Universal Robots URScript: test_first_drawing_6_min3.script

def Machining1():
  # Default parameters:
  global speed_ms = 0.3
  global speed_rads = 0.75
  global accel_mss = 3
  global accel_radss = 1.2
  global blend_radius_m = 0.001

  # Add subprograms here
  # Start of main program
  # Program generated by RoboDK v5.6.5 for UR10e on 02/02/2024 17:04:00
  # Using nominal kinematics.
  blend_radius_m = 0.001
  speed_ms = 1.000
  # set_reference(p[0.133734, -0.230000, -0.014586, 0.000000, 0.000000, 0.000000])
  set_tcp(p[0.000000, 0.000000, 0.252000, 0.000000, 0.000000, 0.000000])
  # Show Tool
  movej([-0.330517, -0.653342, -2.600682, -1.458365, 1.570796, 1.240279],accel_radss,speed_rads,0,blend_radius_m)
  movel([-0.330517, -0.653342, -2.600682, -1.458365, 1.570796, 1.240279],accel_mss,speed_ms,0,blend_radius_m)
  # Splitting Linear movement in 6 (instruction 7: MoveL 3)
  movel([-0.330517, -0.660366, -2.629096, -1.422927, 1.570796, 1.240279],accel_mss,speed_ms,0,blend_radius_m)
  movel([-0.330517, -0.669810, -2.657315, -1.385264, 1.570796, 1.240279],accel_mss,speed_ms,0,blend_radius_m)
  movel([-0.330517, -0.682072, -2.685333, -1.344984, 1.570796, 1.240279],accel_mss,speed_ms,0,blend_radius_m)
  movel([-0.330517, -0.697642, -2.713136, -1.301610, 1.570796, 1.240279],accel_mss,speed_ms,0,blend_radius_m)
  movel([-0.330517, -0.717128, -2.740708, -1.254553, 1.570796, 1.240279],accel_mss,speed_ms,0,blend_radius_m)
  movel([-0.330517, -0.741290, -2.768022, -1.203077, 1.570796, 1.240279],accel_mss,speed_ms,0,blend_radius_m)
  movel([-0.330517, -0.741290, -2.768022, -1.203077, 1.570796, 1.240279],accel_mss,speed_ms,0,blend_radius_m)
  speed_ms = 1.000
  movel([-0.330517, -0.741290, -2.768022, -1.203077, 1.570796, 1.240279],accel_mss,speed_ms,0,blend_radius_m)
  movel([-0.330517, -0.741290, -2.768022, -1.203077, 1.570796, 1.240279],accel_mss,speed_ms,0,blend_radius_m)
  movel([-0.330517, -0.741290, -2.768022, -1.203077, 1.570796, 1.240279],accel_mss,speed_ms,0,blend_radius_m)
  speed_ms = 0.005
  movel([-0.330517, -0.712884, -2.735213, -1.264292, 1.570796, 1.240279],accel_mss,speed_ms,0,blend_radius_m)
  speed_ms = 1.000
  movel([-0.330517, -0.741290, -2.768022, -1.203077, 1.570796, 1.240279],accel_mss,speed_ms,0,blend_radius_m)
  speed_ms = 0.040
  movel([-0.330517, -0.741290, -2.768022, -1.203077, 1.570796, 1.240279],accel_mss,speed_ms,0,blend_radius_m)
  speed_ms = 1.000
  movel([-0.330517, -0.741290, -2.768022, -1.203077, 1.570796, 1.240279],accel_mss,speed_ms,0,blend_radius_m)
  # Splitting Linear movement in 8 (instruction 21: MoveL 12)
  movel([-0.265752, -0.731554, -2.769483, -1.211352, 1.570796, 1.305044],accel_mss,speed_ms,0,blend_radius_m)
  movel([-0.203429, -0.726947, -2.770158, -1.215284, 1.570796, 1.367367],accel_mss,speed_ms,0,blend_radius_m)
  movel([-0.144075, -0.727605, -2.770062, -1.214722, 1.570796, 1.426722],accel_mss,speed_ms,0,blend_radius_m)
  movel([-0.088098, -0.733508, -2.769193, -1.209688, 1.570796, 1.482698],accel_mss,speed_ms,0,blend_radius_m)
  movel([-0.035774, -0.744483, -2.767532, -1.200374, 1.570796, 1.535022],accel_mss,speed_ms,0,blend_radius_m)
  movel([0.012756, -0.760216, -2.765046, -1.187127, 1.570796, 1.583552],accel_mss,speed_ms,0,blend_radius_m)
  movel([0.057475, -0.780279, -2.761690, -1.170420, 1.570796, 1.628271],accel_mss,speed_ms,0,blend_radius_m)
  movel([0.098470, -0.804157, -2.757418, -1.150814, 1.570796, 1.669266],accel_mss,speed_ms,0,blend_radius_m)
  speed_ms = 0.005
  # Splitting Linear movement in 2 (instruction 23: MoveL 13)
  movel([0.098470, -0.822970, -2.773223, -1.116195, 1.570796, 1.669266],accel_mss,speed_ms,0,blend_radius_m)
  movel([0.098470, -0.844049, -2.788876, -1.079465, 1.570796, 1.669266],accel_mss,speed_ms,0,blend_radius_m)
  speed_ms = 0.025
  movel([0.094484, -0.854723, -2.786794, -1.070871, 1.570796, 1.665281],accel_mss,speed_ms,0,blend_radius_m)
  movel([0.092287, -0.860085, -2.785724, -1.066579, 1.570796, 1.663083],accel_mss,speed_ms,0,blend_radius_m)
  movel([0.089913, -0.865446, -2.784638, -1.062305, 1.570796, 1.660710],accel_mss,speed_ms,0,blend_radius_m)
  movel([0.087338, -0.870787, -2.783539, -1.058063, 1.570796, 1.658135],accel_mss,speed_ms,0,blend_radius_m)
  movel([0.084536, -0.876091, -2.782431, -1.053867, 1.570796, 1.655333],accel_mss,speed_ms,0,blend_radius_m)
  movel([0.081477, -0.881347, -2.781317, -1.049725, 1.570796, 1.652273],accel_mss,speed_ms,0,blend_radius_m)
  movel([0.078131, -0.886536, -2.780201, -1.045652, 1.570796, 1.648928],accel_mss,speed_ms,0,blend_radius_m)
  movel([0.079373, -0.884268, -2.780691, -1.047431, 1.570796, 1.650169],accel_mss,speed_ms,0,blend_radius_m)
  movel([0.080517, -0.881424, -2.781300, -1.049665, 1.570796, 1.651313],accel_mss,speed_ms,0,blend_radius_m)
  movel([0.081210, -0.878758, -2.781868, -1.051763, 1.570796, 1.652007],accel_mss,speed_ms,0,blend_radius_m)
  movel([0.081271, -0.877738, -2.782084, -1.052567, 1.570796, 1.652068],accel_mss,speed_ms,0,blend_radius_m)
  movel([0.081086, -0.877049, -2.782229, -1.053110, 1.570796, 1.651882],accel_mss,speed_ms,0,blend_radius_m)
  movel([0.080605, -0.876773, -2.782287, -1.053328, 1.570796, 1.651401],accel_mss,speed_ms,0,blend_radius_m)
  movel([0.079917, -0.877004, -2.782239, -1.053146, 1.570796, 1.650713],accel_mss,speed_ms,0,blend_radius_m)
  movel([0.079063, -0.877672, -2.782098, -1.052619, 1.570796, 1.649859],accel_mss,speed_ms,0,blend_radius_m)
  movel([0.078060, -0.878724, -2.781875, -1.051790, 1.570796, 1.648856],accel_mss,speed_ms,0,blend_radius_m)
  movel([0.075754, -0.881706, -2.781240, -1.049443, 1.570796, 1.646551],accel_mss,speed_ms,0,blend_radius_m)
  movel([0.073242, -0.885438, -2.780438, -1.046513, 1.570796, 1.644038],accel_mss,speed_ms,0,blend_radius_m)
  movel([0.068514, -0.893197, -2.778744, -1.040448, 1.570796, 1.639311],accel_mss,speed_ms,0,blend_radius_m)
  movel([0.065663, -0.898125, -2.777648, -1.036615, 1.570796, 1.636460],accel_mss,speed_ms,0,blend_radius_m)
  movel([0.061416, -0.905014, -2.776092, -1.031283, 1.570796, 1.632212],accel_mss,speed_ms,0,blend_radius_m)
  movel([0.059067, -0.908311, -2.775337, -1.028741, 1.570796, 1.629863],accel_mss,speed_ms,0,blend_radius_m)
  movel([0.056470, -0.911402, -2.774622, -1.026365, 1.570796, 1.627267],accel_mss,speed_ms,0,blend_radius_m)
  movel([0.057008, -0.910476, -2.774837, -1.027076, 1.570796, 1.627804],accel_mss,speed_ms,0,blend_radius_m)
  movel([0.057386, -0.909142, -2.775145, -1.028102, 1.570796, 1.628182],accel_mss,speed_ms,0,blend_radius_m)
  movel([0.057710, -0.905854, -2.775900, -1.030635, 1.570796, 1.628506],accel_mss,speed_ms,0,blend_radius_m)
  movel([0.057532, -0.902784, -2.776599, -1.033006, 1.570796, 1.628328],accel_mss,speed_ms,0,blend_radius_m)
  movel([0.057276, -0.901722, -2.776839, -1.033828, 1.570796, 1.628072],accel_mss,speed_ms,0,blend_radius_m)
  movel([0.056930, -0.901189, -2.776960, -1.034240, 1.570796, 1.627726],accel_mss,speed_ms,0,blend_radius_m)
  movel([0.055907, -0.900938, -2.777016, -1.034434, 1.570796, 1.626704],accel_mss,speed_ms,0,blend_radius_m)
  movel([0.054873, -0.901236, -2.776949, -1.034204, 1.570796, 1.625669],accel_mss,speed_ms,0,blend_radius_m)
  movel([0.053834, -0.901971, -2.776783, -1.033635, 1.570796, 1.624631],accel_mss,speed_ms,0,blend_radius_m)
  movel([0.052803, -0.903040, -2.776541, -1.032808, 1.570796, 1.623599],accel_mss,speed_ms,0,blend_radius_m)
  movel([0.050825, -0.905699, -2.775935, -1.030754, 1.570796, 1.621621],accel_mss,speed_ms,0,blend_radius_m)
  movel([0.049035, -0.908333, -2.775332, -1.028725, 1.570796, 1.619831],accel_mss,speed_ms,0,blend_radius_m)
  movel([0.046096, -0.912299, -2.774414, -1.025676, 1.570796, 1.616892],accel_mss,speed_ms,0,blend_radius_m)
  movel([0.043104, -0.915920, -2.773567, -1.022901, 1.570796, 1.613900],accel_mss,speed_ms,0,blend_radius_m)
  movel([0.039882, -0.919198, -2.772793, -1.020397, 1.570796, 1.610679],accel_mss,speed_ms,0,blend_radius_m)
  movel([0.036270, -0.922107, -2.772101, -1.018181, 1.570796, 1.607066],accel_mss,speed_ms,0,blend_radius_m)
  movel([0.038295, -0.919089, -2.772819, -1.020481, 1.570796, 1.609092],accel_mss,speed_ms,0,blend_radius_m)
  movel([0.039935, -0.916035, -2.773540, -1.022814, 1.570796, 1.610731],accel_mss,speed_ms,0,blend_radius_m)
  movel([0.040448, -0.914524, -2.773894, -1.023970, 1.570796, 1.611244],accel_mss,speed_ms,0,blend_radius_m)
  movel([0.040644, -0.913156, -2.774214, -1.025019, 1.570796, 1.611440],accel_mss,speed_ms,0,blend_radius_m)
  movel([0.040480, -0.912051, -2.774472, -1.025867, 1.570796, 1.611276],accel_mss,speed_ms,0,blend_radius_m)
  movel([0.039889, -0.911359, -2.774632, -1.026398, 1.570796, 1.610686],accel_mss,speed_ms,0,blend_radius_m)
  movel([0.038611, -0.911233, -2.774661, -1.026494, 1.570796, 1.609407],accel_mss,speed_ms,0,blend_radius_m)
  movel([0.036998, -0.911807, -2.774528, -1.026054, 1.570796, 1.607794],accel_mss,speed_ms,0,blend_radius_m)
  movel([0.035210, -0.912847, -2.774286, -1.025256, 1.570796, 1.606006],accel_mss,speed_ms,0,blend_radius_m)
  movel([0.033415, -0.914098, -2.773994, -1.024297, 1.570796, 1.604211],accel_mss,speed_ms,0,blend_radius_m)
  speed_ms = 0.005
  movel([0.033415, -0.904846, -2.767990, -1.039553, 1.570796, 1.604211],accel_mss,speed_ms,0,blend_radius_m)
  speed_ms = 0.040
  movel([0.037572, -0.937768, -2.760014, -1.014607, 1.570796, 1.608368],accel_mss,speed_ms,0,blend_radius_m)
  speed_ms = 0.005
  movel([0.037572, -0.947209, -2.765896, -0.999284, 1.570796, 1.608368],accel_mss,speed_ms,0,blend_radius_m)
  speed_ms = 0.025
  movel([0.038407, -0.944754, -2.766522, -1.001114, 1.570796, 1.609204],accel_mss,speed_ms,0,blend_radius_m)
  movel([0.039504, -0.942229, -2.767161, -1.003000, 1.570796, 1.610300],accel_mss,speed_ms,0,blend_radius_m)
  movel([0.040832, -0.939678, -2.767802, -1.004909, 1.570796, 1.611628],accel_mss,speed_ms,0,blend_radius_m)
  movel([0.042377, -0.937132, -2.768437, -1.006820, 1.570796, 1.613173],accel_mss,speed_ms,0,blend_radius_m)
  movel([0.044112, -0.934624, -2.769059, -1.008705, 1.570796, 1.614908],accel_mss,speed_ms,0,blend_radius_m)
  movel([0.046017, -0.932198, -2.769657, -1.010534, 1.570796, 1.616813],accel_mss,speed_ms,0,blend_radius_m)
  movel([0.048065, -0.929889, -2.770222, -1.012278, 1.570796, 1.618862],accel_mss,speed_ms,0,blend_radius_m)
  movel([0.050239, -0.927730, -2.770747, -1.013912, 1.570796, 1.621035],accel_mss,speed_ms,0,blend_radius_m)
  movel([0.053602, -0.924863, -2.771440, -1.016085, 1.570796, 1.624398],accel_mss,speed_ms,0,blend_radius_m)
  movel([0.056890, -0.922568, -2.771991, -1.017830, 1.570796, 1.627686],accel_mss,speed_ms,0,blend_radius_m)
  movel([0.060092, -0.920808, -2.772411, -1.019170, 1.570796, 1.630888],accel_mss,speed_ms,0,blend_radius_m)
  movel([0.063188, -0.919551, -2.772710, -1.020128, 1.570796, 1.633984],accel_mss,speed_ms,0,blend_radius_m)
  movel([0.066168, -0.918764, -2.772896, -1.020728, 1.570796, 1.636964],accel_mss,speed_ms,0,blend_radius_m)
  movel([0.069022, -0.918410, -2.772980, -1.020999, 1.570796, 1.639818],accel_mss,speed_ms,0,blend_radius_m)
  movel([0.071734, -0.918455, -2.772969, -1.020964, 1.570796, 1.642530],accel_mss,speed_ms,0,blend_radius_m)
  movel([0.074296, -0.918858, -2.772874, -1.020657, 1.570796, 1.645092],accel_mss,speed_ms,0,blend_radius_m)
  movel([0.076697, -0.919580, -2.772703, -1.020106, 1.570796, 1.647493],accel_mss,speed_ms,0,blend_radius_m)
  movel([0.078931, -0.920582, -2.772465, -1.019342, 1.570796, 1.649727],accel_mss,speed_ms,0,blend_radius_m)
  movel([0.082865, -0.923258, -2.771826, -1.017305, 1.570796, 1.653661],accel_mss,speed_ms,0,blend_radius_m)
  movel([0.086044, -0.926549, -2.771034, -1.014807, 1.570796, 1.656840],accel_mss,speed_ms,0,blend_radius_m)
  movel([0.088410, -0.930137, -2.770162, -1.012091, 1.570796, 1.659206],accel_mss,speed_ms,0,blend_radius_m)
  movel([0.090331, -0.934334, -2.769131, -1.008924, 1.570796, 1.661127],accel_mss,speed_ms,0,blend_radius_m)
  movel([0.091833, -0.938890, -2.767999, -1.005500, 1.570796, 1.662629],accel_mss,speed_ms,0,blend_radius_m)
  movel([0.092966, -0.943743, -2.766778, -1.001868, 1.570796, 1.663762],accel_mss,speed_ms,0,blend_radius_m)
  movel([0.093774, -0.948837, -2.765479, -0.998073, 1.570796, 1.664570],accel_mss,speed_ms,0,blend_radius_m)
  movel([0.094306, -0.954114, -2.764115, -0.994160, 1.570796, 1.665103],accel_mss,speed_ms,0,blend_radius_m)
  movel([0.094614, -0.959519, -2.762698, -0.990172, 1.570796, 1.665411],accel_mss,speed_ms,0,blend_radius_m)
  movel([0.094736, -0.970498, -2.759758, -0.982134, 1.570796, 1.665532],accel_mss,speed_ms,0,blend_radius_m)
  movel([0.094750, -0.978142, -2.757660, -0.976588, 1.570796, 1.665546],accel_mss,speed_ms,0,blend_radius_m)
  movel([0.095064, -0.981718, -2.756664, -0.974008, 1.570796, 1.665861],accel_mss,speed_ms,0,blend_radius_m)
  movel([0.095787, -0.984974, -2.755749, -0.971666, 1.570796, 1.666583],accel_mss,speed_ms,0,blend_radius_m)
  movel([0.097346, -0.988765, -2.754674, -0.968950, 1.570796, 1.668143],accel_mss,speed_ms,0,blend_radius_m)
  movel([0.098905, -0.992565, -2.753586, -0.966239, 1.570796, 1.669701],accel_mss,speed_ms,0,blend_radius_m)
  movel([0.099406, -0.994605, -2.752997, -0.964786, 1.570796, 1.670202],accel_mss,speed_ms,0,blend_radius_m)
  movel([0.099571, -0.996815, -2.752356, -0.963218, 1.570796, 1.670367],accel_mss,speed_ms,0,blend_radius_m)
  movel([0.099295, -0.999238, -2.751649, -0.961502, 1.570796, 1.670091],accel_mss,speed_ms,0,blend_radius_m)
  movel([0.098473, -1.001932, -2.750858, -0.959599, 1.570796, 1.669269],accel_mss,speed_ms,0,blend_radius_m)
  movel([0.101094, -0.995138, -2.752843, -0.964408, 1.570796, 1.671890],accel_mss,speed_ms,0,blend_radius_m)
  movel([0.103419, -0.988390, -2.754781, -0.969218, 1.570796, 1.674215],accel_mss,speed_ms,0,blend_radius_m)
  movel([0.107547, -0.974853, -2.758567, -0.978969, 1.570796, 1.678343],accel_mss,speed_ms,0,blend_radius_m)
  movel([0.109649, -0.967278, -2.760629, -0.984483, 1.570796, 1.680446],accel_mss,speed_ms,0,blend_radius_m)
  movel([0.111578, -0.959701, -2.762650, -0.990038, 1.570796, 1.682375],accel_mss,speed_ms,0,blend_radius_m)
  movel([0.115043, -0.944492, -2.766588, -1.001309, 1.570796, 1.685839],accel_mss,speed_ms,0,blend_radius_m)
  movel([0.118016, -0.929526, -2.770310, -1.012552, 1.570796, 1.688812],accel_mss,speed_ms,0,blend_radius_m)
  movel([0.119175, -0.922087, -2.772106, -1.018196, 1.570796, 1.689972],accel_mss,speed_ms,0,blend_radius_m)
  movel([0.119952, -0.914849, -2.773819, -1.023722, 1.570796, 1.690749],accel_mss,speed_ms,0,blend_radius_m)
  movel([0.120167, -0.909356, -2.775096, -1.027937, 1.570796, 1.690963],accel_mss,speed_ms,0,blend_radius_m)
  movel([0.120127, -0.903974, -2.776329, -1.032086, 1.570796, 1.690923],accel_mss,speed_ms,0,blend_radius_m)
  movel([0.120107, -0.898516, -2.777561, -1.036312, 1.570796, 1.690904],accel_mss,speed_ms,0,blend_radius_m)
  movel([0.120387, -0.892798, -2.778832, -1.040759, 1.570796, 1.691183],accel_mss,speed_ms,0,blend_radius_m)
  movel([0.120647, -0.891166, -2.779191, -1.042032, 1.570796, 1.691443],accel_mss,speed_ms,0,blend_radius_m)
  movel([0.121203, -0.889395, -2.779579, -1.043416, 1.570796, 1.692000],accel_mss,speed_ms,0,blend_radius_m)
  movel([0.122110, -0.887725, -2.779942, -1.044721, 1.570796, 1.692906],accel_mss,speed_ms,0,blend_radius_m)
  movel([0.122719, -0.886996, -2.780101, -1.045292, 1.570796, 1.693515],accel_mss,speed_ms,0,blend_radius_m)
  movel([0.123441, -0.886373, -2.780236, -1.045780, 1.570796, 1.694238],accel_mss,speed_ms,0,blend_radius_m)
  movel([0.124465, -0.885837, -2.780352, -1.046200, 1.570796, 1.695262],accel_mss,speed_ms,0,blend_radius_m)
  movel([0.125422, -0.885578, -2.780408, -1.046403, 1.570796, 1.696219],accel_mss,speed_ms,0,blend_radius_m)
  movel([0.130425, -0.884866, -2.780562, -1.046961, 1.570796, 1.701221],accel_mss,speed_ms,0,blend_radius_m)
  movel([0.134885, -0.884918, -2.780550, -1.046921, 1.570796, 1.705681],accel_mss,speed_ms,0,blend_radius_m)
  movel([0.138838, -0.885661, -2.780390, -1.046338, 1.570796, 1.709634],accel_mss,speed_ms,0,blend_radius_m)
  movel([0.142320, -0.887047, -2.780090, -1.045253, 1.570796, 1.713117],accel_mss,speed_ms,0,blend_radius_m)
  movel([0.145368, -0.889002, -2.779664, -1.043723, 1.570796, 1.716164],accel_mss,speed_ms,0,blend_radius_m)
  movel([0.148021, -0.891461, -2.779126, -1.041802, 1.570796, 1.718817],accel_mss,speed_ms,0,blend_radius_m)
  movel([0.150317, -0.894361, -2.778486, -1.039542, 1.570796, 1.721113],accel_mss,speed_ms,0,blend_radius_m)
  movel([0.152293, -0.897642, -2.777756, -1.036991, 1.570796, 1.723089],accel_mss,speed_ms,0,blend_radius_m)
  movel([0.153993, -0.901236, -2.776949, -1.034204, 1.570796, 1.724789],accel_mss,speed_ms,0,blend_radius_m)
  movel([0.155459, -0.905078, -2.776077, -1.031233, 1.570796, 1.726255],accel_mss,speed_ms,0,blend_radius_m)
  movel([0.157842, -0.913264, -2.774189, -1.024936, 1.570796, 1.728639],accel_mss,speed_ms,0,blend_radius_m)
  movel([0.161526, -0.930016, -2.770191, -1.012182, 1.570796, 1.732322],accel_mss,speed_ms,0,blend_radius_m)
  movel([0.162250, -0.932503, -2.769582, -1.010304, 1.570796, 1.733046],accel_mss,speed_ms,0,blend_radius_m)
  movel([0.162856, -0.933490, -2.769339, -1.009560, 1.570796, 1.733653],accel_mss,speed_ms,0,blend_radius_m)
  movel([0.163731, -0.934167, -2.769172, -1.009050, 1.570796, 1.734527],accel_mss,speed_ms,0,blend_radius_m)
  movel([0.165528, -0.934431, -2.769107, -1.008851, 1.570796, 1.736325],accel_mss,speed_ms,0,blend_radius_m)
  movel([0.166517, -0.934232, -2.769156, -1.009001, 1.570796, 1.737313],accel_mss,speed_ms,0,blend_radius_m)
  movel([0.167553, -0.933832, -2.769255, -1.009302, 1.570796, 1.738350],accel_mss,speed_ms,0,blend_radius_m)
  movel([0.169715, -0.932531, -2.769575, -1.010283, 1.570796, 1.740512],accel_mss,speed_ms,0,blend_radius_m)
  movel([0.171931, -0.930687, -2.770027, -1.011675, 1.570796, 1.742727],accel_mss,speed_ms,0,blend_radius_m)
  movel([0.174106, -0.928467, -2.770568, -1.013354, 1.570796, 1.744902],accel_mss,speed_ms,0,blend_radius_m)
  movel([0.176150, -0.926035, -2.771158, -1.015196, 1.570796, 1.746946],accel_mss,speed_ms,0,blend_radius_m)
  movel([0.177974, -0.923550, -2.771756, -1.017083, 1.570796, 1.748770],accel_mss,speed_ms,0,blend_radius_m)
  movel([0.179471, -0.921186, -2.772321, -1.018882, 1.570796, 1.750268],accel_mss,speed_ms,0,blend_radius_m)
  movel([0.181767, -0.917101, -2.773289, -1.021999, 1.570796, 1.752563],accel_mss,speed_ms,0,blend_radius_m)
  movel([0.183931, -0.912963, -2.774259, -1.025166, 1.570796, 1.754728],accel_mss,speed_ms,0,blend_radius_m)
  movel([0.187846, -0.904601, -2.776186, -1.031602, 1.570796, 1.758643],accel_mss,speed_ms,0,blend_radius_m)
  movel([0.191204, -0.896236, -2.778070, -1.038083, 1.570796, 1.762001],accel_mss,speed_ms,0,blend_radius_m)
  movel([0.193979, -0.888009, -2.779881, -1.044499, 1.570796, 1.764775],accel_mss,speed_ms,0,blend_radius_m)
  movel([0.194923, -0.884932, -2.780547, -1.046910, 1.570796, 1.765719],accel_mss,speed_ms,0,blend_radius_m)
  movel([0.196094, -0.881803, -2.781219, -1.049366, 1.570796, 1.766891],accel_mss,speed_ms,0,blend_radius_m)
  movel([0.196862, -0.880242, -2.781553, -1.050595, 1.570796, 1.767658],accel_mss,speed_ms,0,blend_radius_m)
  movel([0.197803, -0.878682, -2.781884, -1.051823, 1.570796, 1.768600],accel_mss,speed_ms,0,blend_radius_m)
  movel([0.198955, -0.877137, -2.782211, -1.053041, 1.570796, 1.769752],accel_mss,speed_ms,0,blend_radius_m)
  movel([0.200357, -0.875619, -2.782530, -1.054240, 1.570796, 1.771153],accel_mss,speed_ms,0,blend_radius_m)
  movel([0.202401, -0.874021, -2.782866, -1.055502, 1.570796, 1.773197],accel_mss,speed_ms,0,blend_radius_m)
  movel([0.204401, -0.873146, -2.783048, -1.056195, 1.570796, 1.775198],accel_mss,speed_ms,0,blend_radius_m)
  movel([0.206224, -0.872912, -2.783097, -1.056380, 1.570796, 1.777021],accel_mss,speed_ms,0,blend_radius_m)
  movel([0.207752, -0.873225, -2.783032, -1.056132, 1.570796, 1.778548],accel_mss,speed_ms,0,blend_radius_m)
  movel([0.209849, -0.874400, -2.782786, -1.055203, 1.570796, 1.780645],accel_mss,speed_ms,0,blend_radius_m)
  movel([0.211668, -0.875985, -2.782453, -1.053950, 1.570796, 1.782464],accel_mss,speed_ms,0,blend_radius_m)
  movel([0.214678, -0.879827, -2.781641, -1.050921, 1.570796, 1.785474],accel_mss,speed_ms,0,blend_radius_m)
  movel([0.215840, -0.881889, -2.781201, -1.049299, 1.570796, 1.786637],accel_mss,speed_ms,0,blend_radius_m)
  movel([0.216722, -0.884138, -2.780719, -1.047533, 1.570796, 1.787518],accel_mss,speed_ms,0,blend_radius_m)
  movel([0.217344, -0.886552, -2.780197, -1.045640, 1.570796, 1.788140],accel_mss,speed_ms,0,blend_radius_m)
  movel([0.217717, -0.889126, -2.779637, -1.043626, 1.570796, 1.788513],accel_mss,speed_ms,0,blend_radius_m)
  movel([0.217858, -0.891840, -2.779043, -1.041507, 1.570796, 1.788654],accel_mss,speed_ms,0,blend_radius_m)
  movel([0.217499, -0.897650, -2.777755, -1.036985, 1.570796, 1.788295],accel_mss,speed_ms,0,blend_radius_m)
  movel([0.217027, -0.900718, -2.777066, -1.034605, 1.570796, 1.787823],accel_mss,speed_ms,0,blend_radius_m)
  movel([0.215585, -0.907111, -2.775612, -1.029666, 1.570796, 1.786381],accel_mss,speed_ms,0,blend_radius_m)
  movel([0.213564, -0.913772, -2.774070, -1.024547, 1.570796, 1.784360],accel_mss,speed_ms,0,blend_radius_m)
  movel([0.211074, -0.920616, -2.772457, -1.019316, 1.570796, 1.781870],accel_mss,speed_ms,0,blend_radius_m)
  movel([0.208233, -0.927540, -2.770794, -1.014056, 1.570796, 1.779029],accel_mss,speed_ms,0,blend_radius_m)
  movel([0.203631, -0.937649, -2.768309, -1.006432, 1.570796, 1.774427],accel_mss,speed_ms,0,blend_radius_m)
  movel([0.201108, -0.942686, -2.767045, -1.002658, 1.570796, 1.771904],accel_mss,speed_ms,0,blend_radius_m)
  movel([0.198410, -0.947683, -2.765775, -0.998931, 1.570796, 1.769207],accel_mss,speed_ms,0,blend_radius_m)
  movel([0.195524, -0.952609, -2.764506, -0.995274, 1.570796, 1.766320],accel_mss,speed_ms,0,blend_radius_m)
  movel([0.192436, -0.957443, -2.763245, -0.991701, 1.570796, 1.763232],accel_mss,speed_ms,0,blend_radius_m)
  movel([0.189119, -0.962171, -2.761996, -0.988222, 1.570796, 1.759915],accel_mss,speed_ms,0,blend_radius_m)
  movel([0.185564, -0.966763, -2.760768, -0.984859, 1.570796, 1.756360],accel_mss,speed_ms,0,blend_radius_m)
  movel([0.180277, -0.972933, -2.759094, -0.980362, 1.570796, 1.751073],accel_mss,speed_ms,0,blend_radius_m)
  movel([0.177371, -0.976017, -2.758247, -0.978125, 1.570796, 1.748167],accel_mss,speed_ms,0,blend_radius_m)
  movel([0.174357, -0.978933, -2.757440, -0.976016, 1.570796, 1.745154],accel_mss,speed_ms,0,blend_radius_m)
  movel([0.171294, -0.981554, -2.756709, -0.974125, 1.570796, 1.742090],accel_mss,speed_ms,0,blend_radius_m)
  movel([0.168232, -0.983759, -2.756091, -0.972539, 1.570796, 1.739028],accel_mss,speed_ms,0,blend_radius_m)
  movel([0.165220, -0.985423, -2.755622, -0.971344, 1.570796, 1.736016],accel_mss,speed_ms,0,blend_radius_m)
  movel([0.163750, -0.986017, -2.755454, -0.970918, 1.570796, 1.734546],accel_mss,speed_ms,0,blend_radius_m)
  movel([0.162314, -0.986425, -2.755338, -0.970625, 1.570796, 1.733110],accel_mss,speed_ms,0,blend_radius_m)
  movel([0.160767, -0.986649, -2.755275, -0.970465, 1.570796, 1.731564],accel_mss,speed_ms,0,blend_radius_m)
  movel([0.159366, -0.986614, -2.755285, -0.970490, 1.570796, 1.730163],accel_mss,speed_ms,0,blend_radius_m)
  movel([0.158098, -0.986347, -2.755361, -0.970681, 1.570796, 1.728894],accel_mss,speed_ms,0,blend_radius_m)
  movel([0.156956, -0.985865, -2.755497, -0.971027, 1.570796, 1.727752],accel_mss,speed_ms,0,blend_radius_m)
  movel([0.155007, -0.984363, -2.755921, -0.972105, 1.570796, 1.725804],accel_mss,speed_ms,0,blend_radius_m)
  movel([0.153455, -0.982282, -2.756506, -0.973601, 1.570796, 1.724251],accel_mss,speed_ms,0,blend_radius_m)
  movel([0.152226, -0.979811, -2.757196, -0.975382, 1.570796, 1.723022],accel_mss,speed_ms,0,blend_radius_m)
  movel([0.151254, -0.977132, -2.757939, -0.977318, 1.570796, 1.722051],accel_mss,speed_ms,0,blend_radius_m)
  movel([0.149812, -0.971891, -2.759378, -0.981119, 1.570796, 1.720608],accel_mss,speed_ms,0,blend_radius_m)
  movel([0.149169, -0.969423, -2.760049, -0.982917, 1.570796, 1.719965],accel_mss,speed_ms,0,blend_radius_m)
  movel([0.148254, -0.967214, -2.760646, -0.984529, 1.570796, 1.719050],accel_mss,speed_ms,0,blend_radius_m)
  movel([0.147575, -0.966367, -2.760874, -0.985148, 1.570796, 1.718371],accel_mss,speed_ms,0,blend_radius_m)
  movel([0.146683, -0.965776, -2.761033, -0.985580, 1.570796, 1.717479],accel_mss,speed_ms,0,blend_radius_m)
  movel([0.145535, -0.965507, -2.761105, -0.985777, 1.570796, 1.716332],accel_mss,speed_ms,0,blend_radius_m)
  movel([0.144083, -0.965620, -2.761075, -0.985695, 1.570796, 1.714879],accel_mss,speed_ms,0,blend_radius_m)
  movel([0.144394, -0.965665, -2.761062, -0.985661, 1.570796, 1.715191],accel_mss,speed_ms,0,blend_radius_m)
  movel([0.144561, -0.965948, -2.760987, -0.985455, 1.570796, 1.715357],accel_mss,speed_ms,0,blend_radius_m)
  movel([0.144480, -0.967165, -2.760659, -0.984565, 1.570796, 1.715276],accel_mss,speed_ms,0,blend_radius_m)
  movel([0.143903, -0.969150, -2.760123, -0.983116, 1.570796, 1.714700],accel_mss,speed_ms,0,blend_radius_m)
  movel([0.142911, -0.971777, -2.759409, -0.981202, 1.570796, 1.713708],accel_mss,speed_ms,0,blend_radius_m)
  movel([0.139967, -0.978457, -2.757572, -0.976360, 1.570796, 1.710763],accel_mss,speed_ms,0,blend_radius_m)
  movel([0.136215, -0.986216, -2.755398, -0.970775, 1.570796, 1.707011],accel_mss,speed_ms,0,blend_radius_m)
  movel([0.128486, -1.001224, -2.751066, -0.960099, 1.570796, 1.699282],accel_mss,speed_ms,0,blend_radius_m)
  movel([0.123866, -1.009671, -2.748554, -0.954164, 1.570796, 1.694663],accel_mss,speed_ms,0,blend_radius_m)
  movel([0.118500, -1.018327, -2.745923, -0.948139, 1.570796, 1.689296],accel_mss,speed_ms,0,blend_radius_m)
  movel([0.113088, -1.026753, -2.743306, -0.942330, 1.570796, 1.683885],accel_mss,speed_ms,0,blend_radius_m)
  movel([0.107607, -1.035034, -2.740679, -0.936676, 1.570796, 1.678403],accel_mss,speed_ms,0,blend_radius_m)
  movel([0.096784, -1.050774, -2.735533, -0.926082, 1.570796, 1.667580],accel_mss,speed_ms,0,blend_radius_m)
  movel([0.091340, -1.058086, -2.733073, -0.921230, 1.570796, 1.662136],accel_mss,speed_ms,0,blend_radius_m)
  movel([0.088492, -1.061586, -2.731879, -0.918923, 1.570796, 1.659288],accel_mss,speed_ms,0,blend_radius_m)
  movel([0.085541, -1.064945, -2.730724, -0.916720, 1.570796, 1.656337],accel_mss,speed_ms,0,blend_radius_m)
  movel([0.082458, -1.068132, -2.729619, -0.914638, 1.570796, 1.653255],accel_mss,speed_ms,0,blend_radius_m)
  movel([0.079236, -1.071121, -2.728575, -0.912693, 1.570796, 1.650032],accel_mss,speed_ms,0,blend_radius_m)
  movel([0.080076, -1.065112, -2.730666, -0.916611, 1.570796, 1.650872],accel_mss,speed_ms,0,blend_radius_m)
  movel([0.080087, -1.063439, -2.731243, -0.917707, 1.570796, 1.650884],accel_mss,speed_ms,0,blend_radius_m)
  movel([0.079804, -1.062865, -2.731441, -0.918083, 1.570796, 1.650600],accel_mss,speed_ms,0,blend_radius_m)
  movel([0.079211, -1.062662, -2.731510, -0.918217, 1.570796, 1.650008],accel_mss,speed_ms,0,blend_radius_m)
  movel([0.078545, -1.062842, -2.731448, -0.918098, 1.570796, 1.649341],accel_mss,speed_ms,0,blend_radius_m)
  movel([0.077831, -1.063265, -2.731303, -0.917821, 1.570796, 1.648627],accel_mss,speed_ms,0,blend_radius_m)
  movel([0.074420, -1.065952, -2.730376, -0.916061, 1.570796, 1.645216],accel_mss,speed_ms,0,blend_radius_m)
  movel([0.072411, -1.067208, -2.729940, -0.915240, 1.570796, 1.643207],accel_mss,speed_ms,0,blend_radius_m)
  movel([0.070406, -1.068179, -2.729603, -0.914607, 1.570796, 1.641202],accel_mss,speed_ms,0,blend_radius_m)
  movel([0.068457, -1.068840, -2.729373, -0.914177, 1.570796, 1.639253],accel_mss,speed_ms,0,blend_radius_m)
  movel([0.067876, -1.068872, -2.729362, -0.914156, 1.570796, 1.638673],accel_mss,speed_ms,0,blend_radius_m)
  movel([0.067717, -1.068534, -2.729479, -0.914376, 1.570796, 1.638514],accel_mss,speed_ms,0,blend_radius_m)
  movel([0.068293, -1.066726, -2.730108, -0.915556, 1.570796, 1.639089],accel_mss,speed_ms,0,blend_radius_m)
  movel([0.068248, -1.066203, -2.730289, -0.915897, 1.570796, 1.639044],accel_mss,speed_ms,0,blend_radius_m)
  movel([0.067937, -1.065895, -2.730396, -0.916098, 1.570796, 1.638733],accel_mss,speed_ms,0,blend_radius_m)
  movel([0.067444, -1.065799, -2.730429, -0.916161, 1.570796, 1.638240],accel_mss,speed_ms,0,blend_radius_m)
  movel([0.066848, -1.065914, -2.730389, -0.916086, 1.570796, 1.637644],accel_mss,speed_ms,0,blend_radius_m)
  movel([0.065582, -1.066611, -2.730147, -0.915630, 1.570796, 1.636378],accel_mss,speed_ms,0,blend_radius_m)
  movel([0.056656, -1.073921, -2.727590, -0.910878, 1.570796, 1.627452],accel_mss,speed_ms,0,blend_radius_m)
  movel([0.059293, -1.071284, -2.728518, -0.912587, 1.570796, 1.630089],accel_mss,speed_ms,0,blend_radius_m)
  movel([0.061894, -1.068447, -2.729509, -0.914432, 1.570796, 1.632691],accel_mss,speed_ms,0,blend_radius_m)
  movel([0.064438, -1.065460, -2.730546, -0.916383, 1.570796, 1.635234],accel_mss,speed_ms,0,blend_radius_m)
  movel([0.066915, -1.062353, -2.731616, -0.918420, 1.570796, 1.637712],accel_mss,speed_ms,0,blend_radius_m)
  movel([0.071603, -1.055938, -2.733800, -0.922651, 1.570796, 1.642399],accel_mss,speed_ms,0,blend_radius_m)
  movel([0.075821, -1.049533, -2.735946, -0.926910, 1.570796, 1.646617],accel_mss,speed_ms,0,blend_radius_m)
  movel([0.080132, -1.042497, -2.738264, -0.931628, 1.570796, 1.650928],accel_mss,speed_ms,0,blend_radius_m)
  movel([0.084250, -1.035307, -2.740592, -0.936491, 1.570796, 1.655047],accel_mss,speed_ms,0,blend_radius_m)
  movel([0.086168, -1.031673, -2.741752, -0.938964, 1.570796, 1.656965],accel_mss,speed_ms,0,blend_radius_m)
  movel([0.087963, -1.028024, -2.742906, -0.941459, 1.570796, 1.658760],accel_mss,speed_ms,0,blend_radius_m)
  movel([0.089601, -1.024373, -2.744051, -0.943965, 1.570796, 1.660397],accel_mss,speed_ms,0,blend_radius_m)
  movel([0.091057, -1.020720, -2.745186, -0.946484, 1.570796, 1.661853],accel_mss,speed_ms,0,blend_radius_m)
  movel([0.091816, -1.018466, -2.745881, -0.948043, 1.570796, 1.662613],accel_mss,speed_ms,0,blend_radius_m)
  movel([0.092410, -1.016236, -2.746564, -0.949589, 1.570796, 1.663206],accel_mss,speed_ms,0,blend_radius_m)
  movel([0.093141, -1.011873, -2.747890, -0.952626, 1.570796, 1.663937],accel_mss,speed_ms,0,blend_radius_m)
  movel([0.093305, -1.007688, -2.749149, -0.955552, 1.570796, 1.664101],accel_mss,speed_ms,0,blend_radius_m)
  movel([0.092955, -1.003734, -2.750326, -0.958330, 1.570796, 1.663751],accel_mss,speed_ms,0,blend_radius_m)
  movel([0.092159, -1.000057, -2.751409, -0.960923, 1.570796, 1.662955],accel_mss,speed_ms,0,blend_radius_m)
  movel([0.090980, -0.996711, -2.752386, -0.963291, 1.570796, 1.661776],accel_mss,speed_ms,0,blend_radius_m)
  movel([0.089473, -0.993750, -2.753244, -0.965394, 1.570796, 1.660269],accel_mss,speed_ms,0,blend_radius_m)
  movel([0.087711, -0.991220, -2.753972, -0.967197, 1.570796, 1.658507],accel_mss,speed_ms,0,blend_radius_m)
  movel([0.086357, -0.990183, -2.754269, -0.967937, 1.570796, 1.657154],accel_mss,speed_ms,0,blend_radius_m)
  movel([0.084665, -0.989854, -2.754363, -0.968172, 1.570796, 1.655461],accel_mss,speed_ms,0,blend_radius_m)
  movel([0.082738, -0.990177, -2.754271, -0.967941, 1.570796, 1.653534],accel_mss,speed_ms,0,blend_radius_m)
  movel([0.080685, -0.991097, -2.754007, -0.967284, 1.570796, 1.651481],accel_mss,speed_ms,0,blend_radius_m)
  movel([0.078604, -0.992552, -2.753590, -0.966248, 1.570796, 1.649400],accel_mss,speed_ms,0,blend_radius_m)
  movel([0.076600, -0.994484, -2.753032, -0.964873, 1.570796, 1.647396],accel_mss,speed_ms,0,blend_radius_m)
  movel([0.074785, -0.996824, -2.752353, -0.963211, 1.570796, 1.645582],accel_mss,speed_ms,0,blend_radius_m)
  movel([0.073255, -0.999514, -2.751568, -0.961307, 1.570796, 1.644052],accel_mss,speed_ms,0,blend_radius_m)
  movel([0.071220, -1.003632, -2.750356, -0.958401, 1.570796, 1.642016],accel_mss,speed_ms,0,blend_radius_m)
  movel([0.069032, -1.007704, -2.749144, -0.955541, 1.570796, 1.639828],accel_mss,speed_ms,0,blend_radius_m)
  movel([0.066672, -1.011696, -2.747944, -0.952749, 1.570796, 1.637469],accel_mss,speed_ms,0,blend_radius_m)
  movel([0.064115, -1.015582, -2.746764, -0.950043, 1.570796, 1.634912],accel_mss,speed_ms,0,blend_radius_m)
  movel([0.061349, -1.019328, -2.745615, -0.947446, 1.570796, 1.632145],accel_mss,speed_ms,0,blend_radius_m)
  movel([0.058346, -1.022909, -2.744507, -0.944973, 1.570796, 1.629142],accel_mss,speed_ms,0,blend_radius_m)
  movel([0.055086, -1.026301, -2.743448, -0.942640, 1.570796, 1.625883],accel_mss,speed_ms,0,blend_radius_m)
  movel([0.051553, -1.029472, -2.742449, -0.940467, 1.570796, 1.622350],accel_mss,speed_ms,0,blend_radius_m)
  movel([0.049638, -1.030916, -2.741992, -0.939481, 1.570796, 1.620435],accel_mss,speed_ms,0,blend_radius_m)
  movel([0.047695, -1.032135, -2.741605, -0.938649, 1.570796, 1.618491],accel_mss,speed_ms,0,blend_radius_m)
  movel([0.043791, -1.034162, -2.740958, -0.937269, 1.570796, 1.614588],accel_mss,speed_ms,0,blend_radius_m)
  movel([0.040756, -1.035447, -2.740547, -0.936395, 1.570796, 1.611552],accel_mss,speed_ms,0,blend_radius_m)
  movel([0.037886, -1.036300, -2.740273, -0.935817, 1.570796, 1.608683],accel_mss,speed_ms,0,blend_radius_m)
  movel([0.035183, -1.036751, -2.740127, -0.935510, 1.570796, 1.605979],accel_mss,speed_ms,0,blend_radius_m)
  movel([0.032632, -1.036838, -2.740100, -0.935452, 1.570796, 1.603429],accel_mss,speed_ms,0,blend_radius_m)
  movel([0.030229, -1.036596, -2.740177, -0.935616, 1.570796, 1.601025],accel_mss,speed_ms,0,blend_radius_m)
  movel([0.027965, -1.036055, -2.740351, -0.935982, 1.570796, 1.598761],accel_mss,speed_ms,0,blend_radius_m)
  movel([0.025843, -1.035244, -2.740612, -0.936533, 1.570796, 1.596639],accel_mss,speed_ms,0,blend_radius_m)
  movel([0.023853, -1.034199, -2.740946, -0.937243, 1.570796, 1.594650],accel_mss,speed_ms,0,blend_radius_m)
  movel([0.021991, -1.032953, -2.741344, -0.938092, 1.570796, 1.592787],accel_mss,speed_ms,0,blend_radius_m)
  movel([0.020254, -1.031528, -2.741798, -0.939063, 1.570796, 1.591051],accel_mss,speed_ms,0,blend_radius_m)
  movel([0.017143, -1.028289, -2.742823, -0.941277, 1.570796, 1.587940],accel_mss,speed_ms,0,blend_radius_m)
  movel([0.014492, -1.024728, -2.743940, -0.943721, 1.570796, 1.585288],accel_mss,speed_ms,0,blend_radius_m)
  movel([0.012279, -1.021103, -2.745067, -0.946219, 1.570796, 1.583076],accel_mss,speed_ms,0,blend_radius_m)
  movel([0.010780, -1.018158, -2.745975, -0.948256, 1.570796, 1.581576],accel_mss,speed_ms,0,blend_radius_m)
  movel([0.009435, -1.014950, -2.746957, -0.950483, 1.570796, 1.580232],accel_mss,speed_ms,0,blend_radius_m)
  movel([0.008265, -1.011488, -2.748007, -0.952895, 1.570796, 1.579062],accel_mss,speed_ms,0,blend_radius_m)
  movel([0.007306, -1.007785, -2.749120, -0.955485, 1.570796, 1.578102],accel_mss,speed_ms,0,blend_radius_m)
  movel([0.006575, -1.003854, -2.750290, -0.958245, 1.570796, 1.577371],accel_mss,speed_ms,0,blend_radius_m)
  movel([0.006105, -0.999708, -2.751511, -0.961169, 1.570796, 1.576901],accel_mss,speed_ms,0,blend_radius_m)
  movel([0.005928, -0.995356, -2.752780, -0.964253, 1.570796, 1.576724],accel_mss,speed_ms,0,blend_radius_m)
  movel([0.006071, -0.990808, -2.754090, -0.967490, 1.570796, 1.576868],accel_mss,speed_ms,0,blend_radius_m)
  movel([0.006563, -0.986075, -2.755438, -0.970876, 1.570796, 1.577359],accel_mss,speed_ms,0,blend_radius_m)
  movel([0.007436, -0.981176, -2.756815, -0.974398, 1.570796, 1.578232],accel_mss,speed_ms,0,blend_radius_m)
  movel([0.008720, -0.976113, -2.758220, -0.978056, 1.570796, 1.579516],accel_mss,speed_ms,0,blend_radius_m)
  movel([0.010453, -0.970900, -2.759648, -0.981841, 1.570796, 1.581249],accel_mss,speed_ms,0,blend_radius_m)
  movel([0.012661, -0.965554, -2.761092, -0.985742, 1.570796, 1.583458],accel_mss,speed_ms,0,blend_radius_m)
  movel([0.015384, -0.960081, -2.762550, -0.989758, 1.570796, 1.586181],accel_mss,speed_ms,0,blend_radius_m)
  movel([0.018649, -0.954506, -2.764013, -0.993870, 1.570796, 1.589446],accel_mss,speed_ms,0,blend_radius_m)
  movel([0.022491, -0.948840, -2.765478, -0.998070, 1.570796, 1.593287],accel_mss,speed_ms,0,blend_radius_m)
  movel([0.024161, -0.946707, -2.766025, -0.999658, 1.570796, 1.594957],accel_mss,speed_ms,0,blend_radius_m)
  movel([0.025079, -0.945746, -2.766269, -1.000373, 1.570796, 1.595875],accel_mss,speed_ms,0,blend_radius_m)
  movel([0.026054, -0.944941, -2.766474, -1.000974, 1.570796, 1.596851],accel_mss,speed_ms,0,blend_radius_m)
  movel([0.027520, -0.944191, -2.766664, -1.001534, 1.570796, 1.598316],accel_mss,speed_ms,0,blend_radius_m)
  movel([0.028823, -0.944015, -2.766709, -1.001665, 1.570796, 1.599619],accel_mss,speed_ms,0,blend_radius_m)
  movel([0.029911, -0.944313, -2.766634, -1.001443, 1.570796, 1.600707],accel_mss,speed_ms,0,blend_radius_m)
  movel([0.030731, -0.944982, -2.766464, -1.000943, 1.570796, 1.601527],accel_mss,speed_ms,0,blend_radius_m)
  movel([0.031881, -0.947147, -2.765912, -0.999330, 1.570796, 1.602677],accel_mss,speed_ms,0,blend_radius_m)
  movel([0.032501, -0.949827, -2.765225, -0.997337, 1.570796, 1.603297],accel_mss,speed_ms,0,blend_radius_m)
  movel([0.033157, -0.955605, -2.763726, -0.993057, 1.570796, 1.603954],accel_mss,speed_ms,0,blend_radius_m)
  movel([0.033560, -0.956499, -2.763492, -0.992397, 1.570796, 1.604356],accel_mss,speed_ms,0,blend_radius_m)
  movel([0.034009, -0.956535, -2.763483, -0.992371, 1.570796, 1.604805],accel_mss,speed_ms,0,blend_radius_m)
  movel([0.034702, -0.956209, -2.763568, -0.992611, 1.570796, 1.605499],accel_mss,speed_ms,0,blend_radius_m)
  movel([0.035843, -0.953482, -2.764280, -0.994627, 1.570796, 1.606639],accel_mss,speed_ms,0,blend_radius_m)
  movel([0.036834, -0.950728, -2.764993, -0.996668, 1.570796, 1.607630],accel_mss,speed_ms,0,blend_radius_m)
  movel([0.037444, -0.959391, -2.762732, -0.990266, 1.570796, 1.608241],accel_mss,speed_ms,0,blend_radius_m)
  movel([0.038358, -0.967755, -2.760500, -0.984134, 1.570796, 1.609155],accel_mss,speed_ms,0,blend_radius_m)
  movel([0.039568, -0.975819, -2.758301, -0.978268, 1.570796, 1.610365],accel_mss,speed_ms,0,blend_radius_m)
  movel([0.041067, -0.983595, -2.756137, -0.972657, 1.570796, 1.611863],accel_mss,speed_ms,0,blend_radius_m)
  movel([0.041844, -0.986867, -2.755213, -0.970309, 1.570796, 1.612640],accel_mss,speed_ms,0,blend_radius_m)
  movel([0.042968, -0.990029, -2.754313, -0.968047, 1.570796, 1.613764],accel_mss,speed_ms,0,blend_radius_m)
  movel([0.043724, -0.991427, -2.753913, -0.967049, 1.570796, 1.614520],accel_mss,speed_ms,0,blend_radius_m)
  movel([0.044642, -0.992627, -2.753568, -0.966194, 1.570796, 1.615439],accel_mss,speed_ms,0,blend_radius_m)
  movel([0.045753, -0.993571, -2.753296, -0.965522, 1.570796, 1.616549],accel_mss,speed_ms,0,blend_radius_m)
  movel([0.047082, -0.994197, -2.753115, -0.965077, 1.570796, 1.617878],accel_mss,speed_ms,0,blend_radius_m)
  movel([0.048145, -0.994403, -2.753056, -0.964930, 1.570796, 1.618941],accel_mss,speed_ms,0,blend_radius_m)
  movel([0.050510, -0.994181, -2.753120, -0.965088, 1.570796, 1.621306],accel_mss,speed_ms,0,blend_radius_m)
  movel([0.051789, -0.993784, -2.753234, -0.965370, 1.570796, 1.622585],accel_mss,speed_ms,0,blend_radius_m)
  movel([0.054481, -0.992511, -2.753601, -0.966277, 1.570796, 1.625277],accel_mss,speed_ms,0,blend_radius_m)
  movel([0.057280, -0.990692, -2.754123, -0.967574, 1.570796, 1.628077],accel_mss,speed_ms,0,blend_radius_m)
  movel([0.060093, -0.988465, -2.754759, -0.969165, 1.570796, 1.630889],accel_mss,speed_ms,0,blend_radius_m)
  movel([0.062827, -0.985950, -2.755473, -0.970966, 1.570796, 1.633623],accel_mss,speed_ms,0,blend_radius_m)
  movel([0.065387, -0.983284, -2.756225, -0.972881, 1.570796, 1.636184],accel_mss,speed_ms,0,blend_radius_m)
  movel([0.067670, -0.980598, -2.756976, -0.974814, 1.570796, 1.638466],accel_mss,speed_ms,0,blend_radius_m)
  speed_ms = 0.005
  movel([0.067670, -0.971009, -2.751222, -0.990158, 1.570796, 1.638466],accel_mss,speed_ms,0,blend_radius_m)
  speed_ms = 0.040
  movel([0.054777, -0.979226, -2.748929, -0.984235, 1.570796, 1.625574],accel_mss,speed_ms,0,blend_radius_m)
  speed_ms = 0.005
  movel([0.054777, -0.988846, -2.754651, -0.968892, 1.570796, 1.625574],accel_mss,speed_ms,0,blend_radius_m)
  speed_ms = 0.025
  movel([0.056594, -0.986607, -2.755287, -0.970495, 1.570796, 1.627391],accel_mss,speed_ms,0,blend_radius_m)
  movel([0.060089, -0.981675, -2.756676, -0.974038, 1.570796, 1.630885],accel_mss,speed_ms,0,blend_radius_m)
  movel([0.061733, -0.979035, -2.757412, -0.975942, 1.570796, 1.632530],accel_mss,speed_ms,0,blend_radius_m)
  movel([0.064740, -0.973541, -2.758927, -0.979920, 1.570796, 1.635536],accel_mss,speed_ms,0,blend_radius_m)
  movel([0.067277, -0.967934, -2.760452, -0.984003, 1.570796, 1.638073],accel_mss,speed_ms,0,blend_radius_m)
  movel([0.068328, -0.965161, -2.761198, -0.986031, 1.570796, 1.639124],accel_mss,speed_ms,0,blend_radius_m)
  movel([0.069210, -0.962440, -2.761924, -0.988025, 1.570796, 1.640006],accel_mss,speed_ms,0,blend_radius_m)
  movel([0.070403, -0.957290, -2.763285, -0.991814, 1.570796, 1.641199],accel_mss,speed_ms,0,blend_radius_m)
  movel([0.070684, -0.954913, -2.763907, -0.993569, 1.570796, 1.641480],accel_mss,speed_ms,0,blend_radius_m)
  movel([0.070726, -0.952718, -2.764478, -0.995193, 1.570796, 1.641522],accel_mss,speed_ms,0,blend_radius_m)
  movel([0.070518, -0.950728, -2.764993, -0.996669, 1.570796, 1.641314],accel_mss,speed_ms,0,blend_radius_m)
  movel([0.070039, -0.948973, -2.765444, -0.997971, 1.570796, 1.640836],accel_mss,speed_ms,0,blend_radius_m)
  movel([0.069145, -0.947071, -2.765932, -0.999387, 1.570796, 1.639941],accel_mss,speed_ms,0,blend_radius_m)
  movel([0.067993, -0.945441, -2.766347, -1.000601, 1.570796, 1.638790],accel_mss,speed_ms,0,blend_radius_m)
  movel([0.066567, -0.944161, -2.766672, -1.001556, 1.570796, 1.637363],accel_mss,speed_ms,0,blend_radius_m)
  movel([0.064853, -0.943313, -2.766887, -1.002189, 1.570796, 1.635649],accel_mss,speed_ms,0,blend_radius_m)
  movel([0.062833, -0.942973, -2.766973, -1.002443, 1.570796, 1.633630],accel_mss,speed_ms,0,blend_radius_m)
  movel([0.060502, -0.943220, -2.766910, -1.002259, 1.570796, 1.631299],accel_mss,speed_ms,0,blend_radius_m)
  movel([0.057846, -0.944130, -2.766680, -1.001579, 1.570796, 1.628642],accel_mss,speed_ms,0,blend_radius_m)
  movel([0.054857, -0.945768, -2.766264, -1.000358, 1.570796, 1.625654],accel_mss,speed_ms,0,blend_radius_m)
  movel([0.052795, -0.947270, -2.765881, -0.999238, 1.570796, 1.623592],accel_mss,speed_ms,0,blend_radius_m)
  movel([0.050789, -0.949066, -2.765420, -0.997903, 1.570796, 1.621585],accel_mss,speed_ms,0,blend_radius_m)
  movel([0.048907, -0.951077, -2.764903, -0.996410, 1.570796, 1.619703],accel_mss,speed_ms,0,blend_radius_m)
  movel([0.047206, -0.953234, -2.764344, -0.994811, 1.570796, 1.618002],accel_mss,speed_ms,0,blend_radius_m)
  movel([0.045744, -0.955466, -2.763763, -0.993161, 1.570796, 1.616540],accel_mss,speed_ms,0,blend_radius_m)
  movel([0.044580, -0.957703, -2.763177, -0.991510, 1.570796, 1.615376],accel_mss,speed_ms,0,blend_radius_m)
  movel([0.043774, -0.959874, -2.762605, -0.989910, 1.570796, 1.614571],accel_mss,speed_ms,0,blend_radius_m)
  movel([0.043376, -0.961917, -2.762063, -0.988409, 1.570796, 1.614172],accel_mss,speed_ms,0,blend_radius_m)
  speed_ms = 0.005
  movel([0.043376, -0.952406, -2.756236, -1.003746, 1.570796, 1.614172],accel_mss,speed_ms,0,blend_radius_m)
  speed_ms = 0.040
  # Splitting Linear movement in 2 (instruction 399: MoveL 378)
  movel([0.095251, -0.959106, -2.754458, -0.998825, 1.570796, 1.666048],accel_mss,speed_ms,0,blend_radius_m)
  movel([0.144369, -0.969768, -2.751564, -0.991057, 1.570796, 1.715166],accel_mss,speed_ms,0,blend_radius_m)
  speed_ms = 0.005
  movel([0.144369, -0.979353, -2.757323, -0.975713, 1.570796, 1.715166],accel_mss,speed_ms,0,blend_radius_m)
  speed_ms = 0.025
  movel([0.142576, -0.989915, -2.754346, -0.968128, 1.570796, 1.713373],accel_mss,speed_ms,0,blend_radius_m)
  movel([0.141323, -0.995271, -2.752804, -0.964313, 1.570796, 1.712119],accel_mss,speed_ms,0,blend_radius_m)
  movel([0.140478, -0.998037, -2.752000, -0.962352, 1.570796, 1.711274],accel_mss,speed_ms,0,blend_radius_m)
  movel([0.139439, -1.000881, -2.751167, -0.960341, 1.570796, 1.710235],accel_mss,speed_ms,0,blend_radius_m)
  movel([0.138085, -1.003939, -2.750265, -0.958185, 1.570796, 1.708881],accel_mss,speed_ms,0,blend_radius_m)
  movel([0.137248, -1.005453, -2.749815, -0.957120, 1.570796, 1.708044],accel_mss,speed_ms,0,blend_radius_m)
  movel([0.136253, -1.006932, -2.749375, -0.956082, 1.570796, 1.707050],accel_mss,speed_ms,0,blend_radius_m)
  movel([0.136298, -1.004628, -2.750060, -0.957700, 1.570796, 1.707094],accel_mss,speed_ms,0,blend_radius_m)
  movel([0.135952, -1.002580, -2.750667, -0.959143, 1.570796, 1.706749],accel_mss,speed_ms,0,blend_radius_m)
  movel([0.135606, -1.002075, -2.750816, -0.959498, 1.570796, 1.706403],accel_mss,speed_ms,0,blend_radius_m)
  movel([0.135231, -1.002120, -2.750802, -0.959466, 1.570796, 1.706027],accel_mss,speed_ms,0,blend_radius_m)
  movel([0.134795, -1.002369, -2.750729, -0.959291, 1.570796, 1.705592],accel_mss,speed_ms,0,blend_radius_m)
  movel([0.133917, -1.003208, -2.750481, -0.958700, 1.570796, 1.704713],accel_mss,speed_ms,0,blend_radius_m)
  movel([0.132686, -1.004805, -2.750008, -0.957576, 1.570796, 1.703482],accel_mss,speed_ms,0,blend_radius_m)
  movel([0.131708, -1.006404, -2.749532, -0.956453, 1.570796, 1.702505],accel_mss,speed_ms,0,blend_radius_m)
  movel([0.130937, -1.007997, -2.749056, -0.955335, 1.570796, 1.701733],accel_mss,speed_ms,0,blend_radius_m)
  movel([0.130326, -1.009580, -2.748581, -0.954227, 1.570796, 1.701122],accel_mss,speed_ms,0,blend_radius_m)
  movel([0.128511, -1.015817, -2.746692, -0.949880, 1.570796, 1.699307],accel_mss,speed_ms,0,blend_radius_m)
  movel([0.127266, -1.019502, -2.745561, -0.947325, 1.570796, 1.698062],accel_mss,speed_ms,0,blend_radius_m)
  movel([0.125795, -1.023214, -2.744412, -0.944763, 1.570796, 1.696591],accel_mss,speed_ms,0,blend_radius_m)
  movel([0.124038, -1.026937, -2.743248, -0.942204, 1.570796, 1.694835],accel_mss,speed_ms,0,blend_radius_m)
  movel([0.121941, -1.030637, -2.742081, -0.939672, 1.570796, 1.692737],accel_mss,speed_ms,0,blend_radius_m)
  movel([0.122563, -1.027876, -2.742953, -0.941560, 1.570796, 1.693359],accel_mss,speed_ms,0,blend_radius_m)
  movel([0.122553, -1.025413, -2.743726, -0.943250, 1.570796, 1.693350],accel_mss,speed_ms,0,blend_radius_m)
  movel([0.122409, -1.024881, -2.743892, -0.943615, 1.570796, 1.693205],accel_mss,speed_ms,0,blend_radius_m)
  movel([0.122040, -1.024589, -2.743984, -0.943817, 1.570796, 1.692837],accel_mss,speed_ms,0,blend_radius_m)
  movel([0.121554, -1.024673, -2.743957, -0.943759, 1.570796, 1.692350],accel_mss,speed_ms,0,blend_radius_m)
  movel([0.121001, -1.025006, -2.743853, -0.943530, 1.570796, 1.691797],accel_mss,speed_ms,0,blend_radius_m)
  movel([0.119921, -1.026062, -2.743523, -0.942804, 1.570796, 1.690717],accel_mss,speed_ms,0,blend_radius_m)
  movel([0.118765, -1.027579, -2.743046, -0.941764, 1.570796, 1.689561],accel_mss,speed_ms,0,blend_radius_m)
  movel([0.117777, -1.029156, -2.742549, -0.940684, 1.570796, 1.688573],accel_mss,speed_ms,0,blend_radius_m)
  movel([0.116176, -1.032397, -2.741521, -0.938471, 1.570796, 1.686972],accel_mss,speed_ms,0,blend_radius_m)
  movel([0.113543, -1.038782, -2.739472, -0.934135, 1.570796, 1.684339],accel_mss,speed_ms,0,blend_radius_m)
  movel([0.111823, -1.042337, -2.738316, -0.931735, 1.570796, 1.682619],accel_mss,speed_ms,0,blend_radius_m)
  movel([0.109889, -1.045870, -2.737158, -0.929361, 1.570796, 1.680686],accel_mss,speed_ms,0,blend_radius_m)
  movel([0.107694, -1.049331, -2.736013, -0.927045, 1.570796, 1.678490],accel_mss,speed_ms,0,blend_radius_m)
  movel([0.105191, -1.052675, -2.734898, -0.924816, 1.570796, 1.675988],accel_mss,speed_ms,0,blend_radius_m)
  movel([0.105698, -1.051155, -2.735406, -0.925828, 1.570796, 1.676494],accel_mss,speed_ms,0,blend_radius_m)
  movel([0.106188, -1.048296, -2.736357, -0.927737, 1.570796, 1.676984],accel_mss,speed_ms,0,blend_radius_m)
  movel([0.106161, -1.046997, -2.736786, -0.928605, 1.570796, 1.676958],accel_mss,speed_ms,0,blend_radius_m)
  movel([0.106006, -1.046488, -2.736954, -0.928947, 1.570796, 1.676802],accel_mss,speed_ms,0,blend_radius_m)
  movel([0.105552, -1.046384, -2.736989, -0.929017, 1.570796, 1.676348],accel_mss,speed_ms,0,blend_radius_m)
  movel([0.104890, -1.046897, -2.736819, -0.928673, 1.570796, 1.675687],accel_mss,speed_ms,0,blend_radius_m)
  movel([0.103405, -1.048535, -2.736277, -0.927577, 1.570796, 1.674202],accel_mss,speed_ms,0,blend_radius_m)
  movel([0.102119, -1.050202, -2.735724, -0.926464, 1.570796, 1.672915],accel_mss,speed_ms,0,blend_radius_m)
  movel([0.099909, -1.053601, -2.734587, -0.924201, 1.570796, 1.670705],accel_mss,speed_ms,0,blend_radius_m)
  movel([0.097790, -1.057030, -2.733431, -0.921928, 1.570796, 1.668586],accel_mss,speed_ms,0,blend_radius_m)
  movel([0.096618, -1.058739, -2.732851, -0.920799, 1.570796, 1.667414],accel_mss,speed_ms,0,blend_radius_m)
  movel([0.095292, -1.060439, -2.732272, -0.919678, 1.570796, 1.666088],accel_mss,speed_ms,0,blend_radius_m)
  movel([0.091838, -1.064374, -2.730921, -0.917094, 1.570796, 1.662635],accel_mss,speed_ms,0,blend_radius_m)
  movel([0.088265, -1.068161, -2.729609, -0.914619, 1.570796, 1.659061],accel_mss,speed_ms,0,blend_radius_m)
  movel([0.084609, -1.071805, -2.728335, -0.912249, 1.570796, 1.655405],accel_mss,speed_ms,0,blend_radius_m)
  movel([0.080897, -1.075327, -2.727092, -0.909969, 1.570796, 1.651693],accel_mss,speed_ms,0,blend_radius_m)
  speed_ms = 0.005
  movel([0.080897, -1.065533, -2.721726, -0.925130, 1.570796, 1.651693],accel_mss,speed_ms,0,blend_radius_m)
  speed_ms = 0.040
  movel([0.052585, -1.037198, -2.731311, -0.943880, 1.570796, 1.623381],accel_mss,speed_ms,0,blend_radius_m)
  speed_ms = 0.005
  movel([0.052585, -1.046964, -2.736797, -0.928628, 1.570796, 1.623381],accel_mss,speed_ms,0,blend_radius_m)
  speed_ms = 0.025
  movel([0.053739, -1.045610, -2.737244, -0.929535, 1.570796, 1.624535],accel_mss,speed_ms,0,blend_radius_m)
  movel([0.054770, -1.044136, -2.737728, -0.930525, 1.570796, 1.625566],accel_mss,speed_ms,0,blend_radius_m)
  movel([0.056627, -1.040964, -2.738764, -0.932661, 1.570796, 1.627423],accel_mss,speed_ms,0,blend_radius_m)
  movel([0.058462, -1.037715, -2.739817, -0.934857, 1.570796, 1.629259],accel_mss,speed_ms,0,blend_radius_m)
  movel([0.059472, -1.036143, -2.740323, -0.935923, 1.570796, 1.630269],accel_mss,speed_ms,0,blend_radius_m)
  movel([0.060595, -1.034655, -2.740800, -0.936934, 1.570796, 1.631391],accel_mss,speed_ms,0,blend_radius_m)
  movel([0.061493, -1.033667, -2.741117, -0.937606, 1.570796, 1.632289],accel_mss,speed_ms,0,blend_radius_m)
  movel([0.062238, -1.033033, -2.741319, -0.938037, 1.570796, 1.633034],accel_mss,speed_ms,0,blend_radius_m)
  movel([0.062844, -1.032714, -2.741420, -0.938254, 1.570796, 1.633640],accel_mss,speed_ms,0,blend_radius_m)
  movel([0.063327, -1.032671, -2.741434, -0.938284, 1.570796, 1.634123],accel_mss,speed_ms,0,blend_radius_m)
  movel([0.063959, -1.033286, -2.741238, -0.937865, 1.570796, 1.634756],accel_mss,speed_ms,0,blend_radius_m)
  movel([0.064238, -1.034579, -2.740825, -0.936985, 1.570796, 1.635035],accel_mss,speed_ms,0,blend_radius_m)
  movel([0.064127, -1.038035, -2.739713, -0.934640, 1.570796, 1.634924],accel_mss,speed_ms,0,blend_radius_m)
  movel([0.063808, -1.040715, -2.738845, -0.932829, 1.570796, 1.634605],accel_mss,speed_ms,0,blend_radius_m)
  movel([0.065855, -1.037473, -2.739895, -0.935021, 1.570796, 1.636651],accel_mss,speed_ms,0,blend_radius_m)
  movel([0.067407, -1.034370, -2.740892, -0.937128, 1.570796, 1.638203],accel_mss,speed_ms,0,blend_radius_m)
  movel([0.068592, -1.031357, -2.741852, -0.939180, 1.570796, 1.639389],accel_mss,speed_ms,0,blend_radius_m)
  movel([0.069527, -1.028402, -2.742787, -0.941200, 1.570796, 1.640323],accel_mss,speed_ms,0,blend_radius_m)
  movel([0.072078, -1.019440, -2.745581, -0.947369, 1.570796, 1.642875],accel_mss,speed_ms,0,blend_radius_m)
  movel([0.073262, -1.016274, -2.746552, -0.949562, 1.570796, 1.644059],accel_mss,speed_ms,0,blend_radius_m)
  movel([0.073925, -1.014982, -2.746947, -0.950460, 1.570796, 1.644722],accel_mss,speed_ms,0,blend_radius_m)
  movel([0.074609, -1.014145, -2.747201, -0.951042, 1.570796, 1.645405],accel_mss,speed_ms,0,blend_radius_m)
  movel([0.075288, -1.013699, -2.747337, -0.951353, 1.570796, 1.646084],accel_mss,speed_ms,0,blend_radius_m)
  movel([0.075933, -1.013587, -2.747371, -0.951431, 1.570796, 1.646729],accel_mss,speed_ms,0,blend_radius_m)
  movel([0.076523, -1.013740, -2.747325, -0.951324, 1.570796, 1.647320],accel_mss,speed_ms,0,blend_radius_m)
  movel([0.077028, -1.014100, -2.747215, -0.951074, 1.570796, 1.647824],accel_mss,speed_ms,0,blend_radius_m)
  movel([0.077688, -1.015177, -2.746887, -0.950325, 1.570796, 1.648484],accel_mss,speed_ms,0,blend_radius_m)
  movel([0.077828, -1.016618, -2.746447, -0.949324, 1.570796, 1.648624],accel_mss,speed_ms,0,blend_radius_m)
  movel([0.077674, -1.018623, -2.745832, -0.947934, 1.570796, 1.648471],accel_mss,speed_ms,0,blend_radius_m)
  movel([0.077147, -1.022419, -2.744659, -0.945311, 1.570796, 1.647943],accel_mss,speed_ms,0,blend_radius_m)
  movel([0.079247, -1.016223, -2.746568, -0.949598, 1.570796, 1.650044],accel_mss,speed_ms,0,blend_radius_m)
  movel([0.080045, -1.013183, -2.747494, -0.951712, 1.570796, 1.650842],accel_mss,speed_ms,0,blend_radius_m)
  movel([0.081117, -1.007272, -2.749273, -0.955844, 1.570796, 1.651913],accel_mss,speed_ms,0,blend_radius_m)
  movel([0.081382, -1.004432, -2.750119, -0.957839, 1.570796, 1.652178],accel_mss,speed_ms,0,blend_radius_m)
  movel([0.081355, -0.999042, -2.751706, -0.961640, 1.570796, 1.652151],accel_mss,speed_ms,0,blend_radius_m)
  speed_ms = 0.005
  movel([0.081355, -0.989388, -2.746025, -0.976977, 1.570796, 1.652151],accel_mss,speed_ms,0,blend_radius_m)
  speed_ms = 0.040
  movel([0.062258, -1.015641, -2.738165, -0.958583, 1.570796, 1.633054],accel_mss,speed_ms,0,blend_radius_m)
  speed_ms = 0.005
  movel([0.062258, -1.025367, -2.743740, -0.943282, 1.570796, 1.633054],accel_mss,speed_ms,0,blend_radius_m)
  speed_ms = 0.025
  movel([0.059858, -1.029084, -2.742572, -0.940733, 1.570796, 1.630654],accel_mss,speed_ms,0,blend_radius_m)
  movel([0.057669, -1.032824, -2.741385, -0.938180, 1.570796, 1.628466],accel_mss,speed_ms,0,blend_radius_m)
  movel([0.053440, -1.040263, -2.738992, -0.933134, 1.570796, 1.624237],accel_mss,speed_ms,0,blend_radius_m)
  movel([0.051127, -1.043941, -2.737792, -0.930656, 1.570796, 1.621923],accel_mss,speed_ms,0,blend_radius_m)
  movel([0.048566, -1.047506, -2.736618, -0.928265, 1.570796, 1.619362],accel_mss,speed_ms,0,blend_radius_m)
  movel([0.045728, -1.050817, -2.735519, -0.926054, 1.570796, 1.616525],accel_mss,speed_ms,0,blend_radius_m)
  movel([0.044200, -1.052333, -2.735012, -0.925044, 1.570796, 1.614997],accel_mss,speed_ms,0,blend_radius_m)
  movel([0.042596, -1.053735, -2.734542, -0.924112, 1.570796, 1.613392],accel_mss,speed_ms,0,blend_radius_m)
  movel([0.043768, -1.052478, -2.734963, -0.924947, 1.570796, 1.614565],accel_mss,speed_ms,0,blend_radius_m)
  movel([0.044992, -1.050668, -2.735568, -0.926153, 1.570796, 1.615788],accel_mss,speed_ms,0,blend_radius_m)
  movel([0.046127, -1.048557, -2.736270, -0.927562, 1.570796, 1.616923],accel_mss,speed_ms,0,blend_radius_m)
  movel([0.047012, -1.046416, -2.736978, -0.928995, 1.570796, 1.617809],accel_mss,speed_ms,0,blend_radius_m)
  movel([0.047502, -1.044502, -2.737608, -0.930279, 1.570796, 1.618298],accel_mss,speed_ms,0,blend_radius_m)
  movel([0.047545, -1.043722, -2.737864, -0.930804, 1.570796, 1.618341],accel_mss,speed_ms,0,blend_radius_m)
  movel([0.047433, -1.043098, -2.738068, -0.931223, 1.570796, 1.618230],accel_mss,speed_ms,0,blend_radius_m)
  movel([0.047146, -1.042665, -2.738210, -0.931515, 1.570796, 1.617942],accel_mss,speed_ms,0,blend_radius_m)
  movel([0.046658, -1.042463, -2.738275, -0.931651, 1.570796, 1.617455],accel_mss,speed_ms,0,blend_radius_m)
  movel([0.045960, -1.042519, -2.738257, -0.931613, 1.570796, 1.616756],accel_mss,speed_ms,0,blend_radius_m)
  movel([0.045023, -1.042871, -2.738142, -0.931376, 1.570796, 1.615819],accel_mss,speed_ms,0,blend_radius_m)
  movel([0.043517, -1.043899, -2.737805, -0.930684, 1.570796, 1.614313],accel_mss,speed_ms,0,blend_radius_m)
  movel([0.037327, -1.049463, -2.735969, -0.926957, 1.570796, 1.608124],accel_mss,speed_ms,0,blend_radius_m)
  movel([0.034681, -1.051571, -2.735267, -0.925551, 1.570796, 1.605478],accel_mss,speed_ms,0,blend_radius_m)
  movel([0.031966, -1.053513, -2.734616, -0.924259, 1.570796, 1.602762],accel_mss,speed_ms,0,blend_radius_m)
  movel([0.029266, -1.055182, -2.734055, -0.923152, 1.570796, 1.600063],accel_mss,speed_ms,0,blend_radius_m)
  movel([0.026666, -1.056459, -2.733624, -0.922306, 1.570796, 1.597462],accel_mss,speed_ms,0,blend_radius_m)
  movel([0.024244, -1.057235, -2.733361, -0.921793, 1.570796, 1.595040],accel_mss,speed_ms,0,blend_radius_m)
  movel([0.022086, -1.057389, -2.733309, -0.921691, 1.570796, 1.592882],accel_mss,speed_ms,0,blend_radius_m)
  movel([0.022777, -1.057232, -2.733363, -0.921795, 1.570796, 1.593573],accel_mss,speed_ms,0,blend_radius_m)
  movel([0.023686, -1.056715, -2.733537, -0.922136, 1.570796, 1.594482],accel_mss,speed_ms,0,blend_radius_m)
  movel([0.025867, -1.054976, -2.734125, -0.923289, 1.570796, 1.596664],accel_mss,speed_ms,0,blend_radius_m)
  movel([0.028010, -1.052908, -2.734820, -0.924661, 1.570796, 1.598806],accel_mss,speed_ms,0,blend_radius_m)
  movel([0.029486, -1.051264, -2.735369, -0.925755, 1.570796, 1.600282],accel_mss,speed_ms,0,blend_radius_m)
  movel([0.030353, -1.050008, -2.735788, -0.926593, 1.570796, 1.601149],accel_mss,speed_ms,0,blend_radius_m)
  movel([0.030677, -1.049179, -2.736064, -0.927146, 1.570796, 1.601473],accel_mss,speed_ms,0,blend_radius_m)
  movel([0.030544, -1.048708, -2.736220, -0.927461, 1.570796, 1.601341],accel_mss,speed_ms,0,blend_radius_m)
  movel([0.030055, -1.048530, -2.736279, -0.927580, 1.570796, 1.600851],accel_mss,speed_ms,0,blend_radius_m)
  movel([0.028394, -1.048778, -2.736197, -0.927414, 1.570796, 1.599190],accel_mss,speed_ms,0,blend_radius_m)
  movel([0.026468, -1.049381, -2.735997, -0.927012, 1.570796, 1.597264],accel_mss,speed_ms,0,blend_radius_m)
  movel([0.022092, -1.050747, -2.735542, -0.926100, 1.570796, 1.592888],accel_mss,speed_ms,0,blend_radius_m)
  movel([0.017739, -1.051735, -2.735212, -0.925442, 1.570796, 1.588535],accel_mss,speed_ms,0,blend_radius_m)
  movel([0.015686, -1.051953, -2.735139, -0.925297, 1.570796, 1.586482],accel_mss,speed_ms,0,blend_radius_m)
  movel([0.013777, -1.051912, -2.735153, -0.925324, 1.570796, 1.584574],accel_mss,speed_ms,0,blend_radius_m)
  movel([0.012060, -1.051556, -2.735272, -0.925561, 1.570796, 1.582856],accel_mss,speed_ms,0,blend_radius_m)
  movel([0.010581, -1.050830, -2.735514, -0.926045, 1.570796, 1.581377],accel_mss,speed_ms,0,blend_radius_m)
  movel([0.013190, -1.049987, -2.735795, -0.926607, 1.570796, 1.583987],accel_mss,speed_ms,0,blend_radius_m)
  movel([0.014621, -1.049217, -2.736051, -0.927121, 1.570796, 1.585417],accel_mss,speed_ms,0,blend_radius_m)
  movel([0.015257, -1.048713, -2.736218, -0.927457, 1.570796, 1.586053],accel_mss,speed_ms,0,blend_radius_m)
  movel([0.015800, -1.048113, -2.736417, -0.927859, 1.570796, 1.586596],accel_mss,speed_ms,0,blend_radius_m)
  movel([0.016023, -1.047656, -2.736569, -0.928165, 1.570796, 1.586820],accel_mss,speed_ms,0,blend_radius_m)
  movel([0.015994, -1.047241, -2.736706, -0.928443, 1.570796, 1.586790],accel_mss,speed_ms,0,blend_radius_m)
  movel([0.015315, -1.046531, -2.736940, -0.928918, 1.570796, 1.586112],accel_mss,speed_ms,0,blend_radius_m)
  movel([0.013996, -1.045971, -2.737125, -0.929293, 1.570796, 1.584792],accel_mss,speed_ms,0,blend_radius_m)
  movel([0.012280, -1.045538, -2.737267, -0.929583, 1.570796, 1.583076],accel_mss,speed_ms,0,blend_radius_m)
  movel([0.006259, -1.044678, -2.737550, -0.930161, 1.570796, 1.577055],accel_mss,speed_ms,0,blend_radius_m)
  movel([0.004079, -1.044014, -2.737768, -0.930607, 1.570796, 1.574875],accel_mss,speed_ms,0,blend_radius_m)
  movel([0.002111, -1.043044, -2.738086, -0.931260, 1.570796, 1.572908],accel_mss,speed_ms,0,blend_radius_m)
  movel([0.000486, -1.041680, -2.738531, -0.932178, 1.570796, 1.571283],accel_mss,speed_ms,0,blend_radius_m)
  movel([-0.000685, -1.039839, -2.739129, -0.933420, 1.570796, 1.570112],accel_mss,speed_ms,0,blend_radius_m)
  movel([0.001330, -1.040574, -2.738891, -0.932924, 1.570796, 1.572126],accel_mss,speed_ms,0,blend_radius_m)
  movel([0.002588, -1.040696, -2.738851, -0.932842, 1.570796, 1.573385],accel_mss,speed_ms,0,blend_radius_m)
  movel([0.003813, -1.040380, -2.738954, -0.933055, 1.570796, 1.574610],accel_mss,speed_ms,0,blend_radius_m)
  movel([0.004986, -1.039551, -2.739223, -0.933615, 1.570796, 1.575782],accel_mss,speed_ms,0,blend_radius_m)
  movel([0.005693, -1.038578, -2.739538, -0.934273, 1.570796, 1.576489],accel_mss,speed_ms,0,blend_radius_m)
  movel([0.005907, -1.037594, -2.739856, -0.934939, 1.570796, 1.576703],accel_mss,speed_ms,0,blend_radius_m)
  movel([0.005604, -1.036725, -2.740136, -0.935528, 1.570796, 1.576400],accel_mss,speed_ms,0,blend_radius_m)
  movel([0.003068, -1.032794, -2.741395, -0.938200, 1.570796, 1.573864],accel_mss,speed_ms,0,blend_radius_m)
  movel([0.001141, -1.028435, -2.742777, -0.941178, 1.570796, 1.571937],accel_mss,speed_ms,0,blend_radius_m)
  movel([0.000453, -1.026021, -2.743536, -0.942833, 1.570796, 1.571250],accel_mss,speed_ms,0,blend_radius_m)
  movel([-0.000030, -1.023414, -2.744350, -0.944625, 1.570796, 1.570766],accel_mss,speed_ms,0,blend_radius_m)
  movel([-0.000289, -1.020581, -2.745228, -0.946579, 1.570796, 1.570507],accel_mss,speed_ms,0,blend_radius_m)
  movel([-0.000305, -1.017494, -2.746179, -0.948716, 1.570796, 1.570491],accel_mss,speed_ms,0,blend_radius_m)
  speed_ms = 0.005
  movel([-0.000305, -1.007787, -2.740571, -0.964031, 1.570796, 1.570491],accel_mss,speed_ms,0,blend_radius_m)
  speed_ms = 0.040
  movel([-0.041269, -1.000189, -2.742854, -0.969346, 1.570796, 1.529527],accel_mss,speed_ms,0,blend_radius_m)
  speed_ms = 0.005
  movel([-0.041269, -1.009876, -2.748493, -0.954021, 1.570796, 1.529527],accel_mss,speed_ms,0,blend_radius_m)
  speed_ms = 0.025
  movel([-0.037935, -1.004303, -2.750157, -0.957929, 1.570796, 1.532862],accel_mss,speed_ms,0,blend_radius_m)
  movel([-0.034722, -0.998672, -2.751815, -0.961902, 1.570796, 1.536074],accel_mss,speed_ms,0,blend_radius_m)
  movel([-0.028597, -0.987207, -2.755117, -0.970065, 1.570796, 1.542199],accel_mss,speed_ms,0,blend_radius_m)
  movel([-0.022885, -0.975503, -2.758389, -0.978498, 1.570796, 1.547912],accel_mss,speed_ms,0,blend_radius_m)
  movel([-0.017602, -0.963598, -2.761616, -0.987176, 1.570796, 1.553194],accel_mss,speed_ms,0,blend_radius_m)
  movel([-0.012765, -0.951528, -2.764786, -0.996075, 1.570796, 1.558032],accel_mss,speed_ms,0,blend_radius_m)
  movel([-0.008393, -0.939340, -2.767886, -1.005162, 1.570796, 1.562403],accel_mss,speed_ms,0,blend_radius_m)
  movel([-0.004507, -0.927088, -2.770903, -1.014398, 1.570796, 1.566289],accel_mss,speed_ms,0,blend_radius_m)
  movel([-0.001128, -0.914816, -2.773826, -1.023747, 1.570796, 1.569668],accel_mss,speed_ms,0,blend_radius_m)
  movel([0.001717, -0.902594, -2.776642, -1.033153, 1.570796, 1.572514],accel_mss,speed_ms,0,blend_radius_m)
  movel([0.004003, -0.890482, -2.779341, -1.042566, 1.570796, 1.574800],accel_mss,speed_ms,0,blend_radius_m)
  movel([0.005699, -0.878552, -2.781912, -1.051926, 1.570796, 1.576495],accel_mss,speed_ms,0,blend_radius_m)
  movel([0.006772, -0.866879, -2.784345, -1.061165, 1.570796, 1.577568],accel_mss,speed_ms,0,blend_radius_m)
  movel([0.007201, -0.855532, -2.786634, -1.070223, 1.570796, 1.577998],accel_mss,speed_ms,0,blend_radius_m)
  movel([0.006944, -0.844605, -2.788769, -1.079015, 1.570796, 1.577741],accel_mss,speed_ms,0,blend_radius_m)
  movel([0.005975, -0.834183, -2.790743, -1.087464, 1.570796, 1.576771],accel_mss,speed_ms,0,blend_radius_m)
  movel([0.003369, -0.819440, -2.793433, -1.099516, 1.570796, 1.574166],accel_mss,speed_ms,0,blend_radius_m)
  movel([0.003313, -0.816685, -2.793923, -1.101781, 1.570796, 1.574110],accel_mss,speed_ms,0,blend_radius_m)
  movel([0.003753, -0.813590, -2.794468, -1.104331, 1.570796, 1.574550],accel_mss,speed_ms,0,blend_radius_m)
  movel([0.005074, -0.808944, -2.795278, -1.108168, 1.570796, 1.575870],accel_mss,speed_ms,0,blend_radius_m)
  movel([0.006722, -0.805081, -2.795942, -1.111366, 1.570796, 1.577519],accel_mss,speed_ms,0,blend_radius_m)
  movel([0.007652, -0.803432, -2.796223, -1.112734, 1.570796, 1.578448],accel_mss,speed_ms,0,blend_radius_m)
  movel([0.009696, -0.800651, -2.796694, -1.115044, 1.570796, 1.580493],accel_mss,speed_ms,0,blend_radius_m)
  movel([0.010791, -0.799517, -2.796885, -1.115987, 1.570796, 1.581587],accel_mss,speed_ms,0,blend_radius_m)
  movel([0.013113, -0.797712, -2.797187, -1.117490, 1.570796, 1.583910],accel_mss,speed_ms,0,blend_radius_m)
  movel([0.015556, -0.796485, -2.797392, -1.118513, 1.570796, 1.586352],accel_mss,speed_ms,0,blend_radius_m)
  movel([0.018066, -0.795782, -2.797509, -1.119099, 1.570796, 1.588863],accel_mss,speed_ms,0,blend_radius_m)
  movel([0.020598, -0.795547, -2.797548, -1.119294, 1.570796, 1.591395],accel_mss,speed_ms,0,blend_radius_m)
  movel([0.023097, -0.795718, -2.797519, -1.119152, 1.570796, 1.593894],accel_mss,speed_ms,0,blend_radius_m)
  movel([0.025518, -0.796238, -2.797433, -1.118718, 1.570796, 1.596315],accel_mss,speed_ms,0,blend_radius_m)
  movel([0.029924, -0.798062, -2.797129, -1.117198, 1.570796, 1.600720],accel_mss,speed_ms,0,blend_radius_m)
  movel([0.033447, -0.800514, -2.796717, -1.115158, 1.570796, 1.604244],accel_mss,speed_ms,0,blend_radius_m)
  movel([0.035752, -0.803047, -2.796288, -1.113054, 1.570796, 1.606548],accel_mss,speed_ms,0,blend_radius_m)
  movel([0.037774, -0.806705, -2.795663, -1.110020, 1.570796, 1.608570],accel_mss,speed_ms,0,blend_radius_m)
  movel([0.039406, -0.810763, -2.794962, -1.106664, 1.570796, 1.610203],accel_mss,speed_ms,0,blend_radius_m)
  movel([0.041880, -0.819628, -2.793400, -1.099362, 1.570796, 1.612676],accel_mss,speed_ms,0,blend_radius_m)
  movel([0.043907, -0.828811, -2.791737, -1.091841, 1.570796, 1.614703],accel_mss,speed_ms,0,blend_radius_m)
  movel([0.046189, -0.837534, -2.790115, -1.084741, 1.570796, 1.616985],accel_mss,speed_ms,0,blend_radius_m)
  movel([0.048787, -0.844777, -2.788736, -1.078877, 1.570796, 1.619584],accel_mss,speed_ms,0,blend_radius_m)
  movel([0.050495, -0.847950, -2.788122, -1.076317, 1.570796, 1.621292],accel_mss,speed_ms,0,blend_radius_m)
  movel([0.052701, -0.850557, -2.787614, -1.074217, 1.570796, 1.623497],accel_mss,speed_ms,0,blend_radius_m)
  movel([0.054025, -0.851416, -2.787446, -1.073527, 1.570796, 1.624822],accel_mss,speed_ms,0,blend_radius_m)
  movel([0.054860, -0.851576, -2.787415, -1.073398, 1.570796, 1.625656],accel_mss,speed_ms,0,blend_radius_m)
  movel([0.055847, -0.851449, -2.787439, -1.073500, 1.570796, 1.626643],accel_mss,speed_ms,0,blend_radius_m)
  movel([0.057282, -0.850808, -2.787565, -1.074016, 1.570796, 1.628078],accel_mss,speed_ms,0,blend_radius_m)
  movel([0.058791, -0.849749, -2.787772, -1.074868, 1.570796, 1.629587],accel_mss,speed_ms,0,blend_radius_m)
  movel([0.061813, -0.846919, -2.788322, -1.077148, 1.570796, 1.632609],accel_mss,speed_ms,0,blend_radius_m)
  movel([0.065119, -0.843315, -2.789016, -1.080058, 1.570796, 1.635915],accel_mss,speed_ms,0,blend_radius_m)
  movel([0.068277, -0.839555, -2.789733, -1.083101, 1.570796, 1.639073],accel_mss,speed_ms,0,blend_radius_m)
  movel([0.074274, -0.831668, -2.791210, -1.089511, 1.570796, 1.645070],accel_mss,speed_ms,0,blend_radius_m)
  movel([0.085956, -0.815233, -2.794179, -1.102977, 1.570796, 1.656752],accel_mss,speed_ms,0,blend_radius_m)
  movel([0.091724, -0.807543, -2.795519, -1.109326, 1.570796, 1.662520],accel_mss,speed_ms,0,blend_radius_m)
  movel([0.095118, -0.803369, -2.796234, -1.112787, 1.570796, 1.665914],accel_mss,speed_ms,0,blend_radius_m)
  movel([0.098550, -0.799589, -2.796872, -1.115927, 1.570796, 1.669346],accel_mss,speed_ms,0,blend_radius_m)
  movel([0.100208, -0.797990, -2.797141, -1.117259, 1.570796, 1.671005],accel_mss,speed_ms,0,blend_radius_m)
  movel([0.101792, -0.796663, -2.797362, -1.118364, 1.570796, 1.672589],accel_mss,speed_ms,0,blend_radius_m)
  movel([0.103267, -0.795668, -2.797528, -1.119194, 1.570796, 1.674063],accel_mss,speed_ms,0,blend_radius_m)
  movel([0.104605, -0.795066, -2.797627, -1.119695, 1.570796, 1.675402],accel_mss,speed_ms,0,blend_radius_m)
  movel([0.105774, -0.794912, -2.797653, -1.119824, 1.570796, 1.676571],accel_mss,speed_ms,0,blend_radius_m)
  movel([0.106748, -0.795260, -2.797595, -1.119533, 1.570796, 1.677544],accel_mss,speed_ms,0,blend_radius_m)
  movel([0.107496, -0.796175, -2.797443, -1.118771, 1.570796, 1.678292],accel_mss,speed_ms,0,blend_radius_m)
  movel([0.107985, -0.797711, -2.797187, -1.117490, 1.570796, 1.678781],accel_mss,speed_ms,0,blend_radius_m)
  movel([0.108380, -0.800826, -2.796664, -1.114899, 1.570796, 1.679177],accel_mss,speed_ms,0,blend_radius_m)
  movel([0.108432, -0.804122, -2.796105, -1.112161, 1.570796, 1.679228],accel_mss,speed_ms,0,blend_radius_m)
  movel([0.108163, -0.807576, -2.795514, -1.109300, 1.570796, 1.678960],accel_mss,speed_ms,0,blend_radius_m)
  movel([0.107597, -0.811173, -2.794891, -1.106325, 1.570796, 1.678393],accel_mss,speed_ms,0,blend_radius_m)
  movel([0.106747, -0.814887, -2.794240, -1.103262, 1.570796, 1.677543],accel_mss,speed_ms,0,blend_radius_m)
  movel([0.105636, -0.818702, -2.793565, -1.100122, 1.570796, 1.676432],accel_mss,speed_ms,0,blend_radius_m)
  movel([0.104281, -0.822601, -2.792866, -1.096922, 1.570796, 1.675078],accel_mss,speed_ms,0,blend_radius_m)
  movel([0.102705, -0.826566, -2.792147, -1.093676, 1.570796, 1.673502],accel_mss,speed_ms,0,blend_radius_m)
  movel([0.098963, -0.834616, -2.790662, -1.087111, 1.570796, 1.669759],accel_mss,speed_ms,0,blend_radius_m)
  movel([0.094548, -0.842729, -2.789128, -1.080531, 1.570796, 1.665345],accel_mss,speed_ms,0,blend_radius_m)
  movel([0.089597, -0.850783, -2.787570, -1.074036, 1.570796, 1.660394],accel_mss,speed_ms,0,blend_radius_m)
  movel([0.084252, -0.858654, -2.786011, -1.067723, 1.570796, 1.655048],accel_mss,speed_ms,0,blend_radius_m)
  movel([0.071998, -0.875774, -2.782498, -1.054117, 1.570796, 1.642794],accel_mss,speed_ms,0,blend_radius_m)
  movel([0.065571, -0.884067, -2.780734, -1.047588, 1.570796, 1.636367],accel_mss,speed_ms,0,blend_radius_m)
  movel([0.062299, -0.887949, -2.779894, -1.044546, 1.570796, 1.633095],accel_mss,speed_ms,0,blend_radius_m)
  movel([0.058990, -0.891585, -2.779099, -1.041705, 1.570796, 1.629786],accel_mss,speed_ms,0,blend_radius_m)
  movel([0.056838, -0.893746, -2.778622, -1.040020, 1.570796, 1.627635],accel_mss,speed_ms,0,blend_radius_m)
  movel([0.054684, -0.895698, -2.778190, -1.038501, 1.570796, 1.625481],accel_mss,speed_ms,0,blend_radius_m)
  movel([0.052541, -0.897410, -2.777808, -1.037171, 1.570796, 1.623337],accel_mss,speed_ms,0,blend_radius_m)
  movel([0.050425, -0.898849, -2.777486, -1.036054, 1.570796, 1.621221],accel_mss,speed_ms,0,blend_radius_m)
  movel([0.048357, -0.899982, -2.777232, -1.035176, 1.570796, 1.619154],accel_mss,speed_ms,0,blend_radius_m)
  movel([0.046350, -0.900779, -2.777052, -1.034558, 1.570796, 1.617147],accel_mss,speed_ms,0,blend_radius_m)
  movel([0.044425, -0.901200, -2.776957, -1.034232, 1.570796, 1.615221],accel_mss,speed_ms,0,blend_radius_m)
  movel([0.042592, -0.901213, -2.776954, -1.034221, 1.570796, 1.613389],accel_mss,speed_ms,0,blend_radius_m)
  movel([0.040937, -0.900784, -2.777051, -1.034554, 1.570796, 1.611733],accel_mss,speed_ms,0,blend_radius_m)
  movel([0.039563, -0.899997, -2.777228, -1.035163, 1.570796, 1.610360],accel_mss,speed_ms,0,blend_radius_m)
  movel([0.034961, -0.895626, -2.778206, -1.038558, 1.570796, 1.605758],accel_mss,speed_ms,0,blend_radius_m)
  movel([0.033548, -0.894829, -2.778383, -1.039178, 1.570796, 1.604344],accel_mss,speed_ms,0,blend_radius_m)
  movel([0.031832, -0.894400, -2.778478, -1.039511, 1.570796, 1.602629],accel_mss,speed_ms,0,blend_radius_m)
  movel([0.031048, -0.894507, -2.778454, -1.039428, 1.570796, 1.601844],accel_mss,speed_ms,0,blend_radius_m)
  movel([0.030681, -0.895011, -2.778342, -1.039036, 1.570796, 1.601477],accel_mss,speed_ms,0,blend_radius_m)
  movel([0.030199, -0.896165, -2.778086, -1.038138, 1.570796, 1.600996],accel_mss,speed_ms,0,blend_radius_m)
  movel([0.028942, -0.900083, -2.777209, -1.035097, 1.570796, 1.599739],accel_mss,speed_ms,0,blend_radius_m)
  movel([0.025811, -0.911762, -2.774539, -1.026089, 1.570796, 1.596608],accel_mss,speed_ms,0,blend_radius_m)
  movel([0.020960, -0.930998, -2.769951, -1.011440, 1.570796, 1.591756],accel_mss,speed_ms,0,blend_radius_m)
  movel([0.017470, -0.941288, -2.767398, -1.003703, 1.570796, 1.588266],accel_mss,speed_ms,0,blend_radius_m)
  movel([0.013608, -0.951543, -2.764782, -0.996064, 1.570796, 1.584404],accel_mss,speed_ms,0,blend_radius_m)
  movel([0.009426, -0.961733, -2.762112, -0.988544, 1.570796, 1.580223],accel_mss,speed_ms,0,blend_radius_m)
  movel([0.004989, -0.971817, -2.759398, -0.981173, 1.570796, 1.575785],accel_mss,speed_ms,0,blend_radius_m)
  movel([-0.000886, -0.984560, -2.755865, -0.971963, 1.570796, 1.569910],accel_mss,speed_ms,0,blend_radius_m)
  movel([-0.006924, -0.997139, -2.752262, -0.962988, 1.570796, 1.563873],accel_mss,speed_ms,0,blend_radius_m)
  movel([-0.013170, -1.009509, -2.748603, -0.954277, 1.570796, 1.557626],accel_mss,speed_ms,0,blend_radius_m)
  movel([-0.019682, -1.021628, -2.744905, -0.945857, 1.570796, 1.551114],accel_mss,speed_ms,0,blend_radius_m)
  movel([-0.026507, -1.033447, -2.741187, -0.937755, 1.570796, 1.544290],accel_mss,speed_ms,0,blend_radius_m)
  movel([-0.030048, -1.039233, -2.739326, -0.933830, 1.570796, 1.540749],accel_mss,speed_ms,0,blend_radius_m)
  movel([-0.033689, -1.044934, -2.737466, -0.929989, 1.570796, 1.537107],accel_mss,speed_ms,0,blend_radius_m)
  movel([-0.037435, -1.050545, -2.735609, -0.926235, 1.570796, 1.533362],accel_mss,speed_ms,0,blend_radius_m)
  movel([-0.041287, -1.056057, -2.733760, -0.922572, 1.570796, 1.529509],accel_mss,speed_ms,0,blend_radius_m)
  movel([-0.045255, -1.061474, -2.731918, -0.918997, 1.570796, 1.525541],accel_mss,speed_ms,0,blend_radius_m)
  movel([-0.049349, -1.066787, -2.730086, -0.915515, 1.570796, 1.521448],accel_mss,speed_ms,0,blend_radius_m)
  movel([-0.054352, -1.072959, -2.727929, -0.911501, 1.570796, 1.516444],accel_mss,speed_ms,0,blend_radius_m)
  movel([-0.056958, -1.075922, -2.726882, -0.909585, 1.570796, 1.513838],accel_mss,speed_ms,0,blend_radius_m)
  movel([-0.061649, -1.080682, -2.725183, -0.906524, 1.570796, 1.509147],accel_mss,speed_ms,0,blend_radius_m)
  movel([-0.064077, -1.082853, -2.724401, -0.905135, 1.570796, 1.506719],accel_mss,speed_ms,0,blend_radius_m)
  movel([-0.066519, -1.084589, -2.723774, -0.904026, 1.570796, 1.504277],accel_mss,speed_ms,0,blend_radius_m)
  movel([-0.067609, -1.085083, -2.723594, -0.903711, 1.570796, 1.503188],accel_mss,speed_ms,0,blend_radius_m)
  movel([-0.068545, -1.085221, -2.723544, -0.903623, 1.570796, 1.502251],accel_mss,speed_ms,0,blend_radius_m)
  movel([-0.067892, -1.082630, -2.724482, -0.905277, 1.570796, 1.502904],accel_mss,speed_ms,0,blend_radius_m)
  movel([-0.067596, -1.080174, -2.725365, -0.906850, 1.570796, 1.503200],accel_mss,speed_ms,0,blend_radius_m)
  movel([-0.067673, -1.079114, -2.725745, -0.907530, 1.570796, 1.503124],accel_mss,speed_ms,0,blend_radius_m)
  movel([-0.067948, -1.078230, -2.726061, -0.908099, 1.570796, 1.502849],accel_mss,speed_ms,0,blend_radius_m)
  movel([-0.068456, -1.077565, -2.726298, -0.908527, 1.570796, 1.502340],accel_mss,speed_ms,0,blend_radius_m)
  movel([-0.069242, -1.077177, -2.726436, -0.908776, 1.570796, 1.501554],accel_mss,speed_ms,0,blend_radius_m)
  movel([-0.071652, -1.076950, -2.726516, -0.908923, 1.570796, 1.499145],accel_mss,speed_ms,0,blend_radius_m)
  movel([-0.072322, -1.076607, -2.726638, -0.909144, 1.570796, 1.498475],accel_mss,speed_ms,0,blend_radius_m)
  movel([-0.072785, -1.076049, -2.726836, -0.909503, 1.570796, 1.498011],accel_mss,speed_ms,0,blend_radius_m)
  movel([-0.073179, -1.074430, -2.727410, -0.910549, 1.570796, 1.497617],accel_mss,speed_ms,0,blend_radius_m)
  movel([-0.073051, -1.072375, -2.728135, -0.911879, 1.570796, 1.497746],accel_mss,speed_ms,0,blend_radius_m)
  movel([-0.072608, -1.070173, -2.728907, -0.913309, 1.570796, 1.498188],accel_mss,speed_ms,0,blend_radius_m)
  movel([-0.070858, -1.063387, -2.731261, -0.917741, 1.570796, 1.499938],accel_mss,speed_ms,0,blend_radius_m)
  movel([-0.068698, -1.056368, -2.733655, -0.922366, 1.570796, 1.502098],accel_mss,speed_ms,0,blend_radius_m)
  movel([-0.067395, -1.052787, -2.734860, -0.924742, 1.570796, 1.503402],accel_mss,speed_ms,0,blend_radius_m)
  movel([-0.065910, -1.049164, -2.736069, -0.927157, 1.570796, 1.504886],accel_mss,speed_ms,0,blend_radius_m)
  movel([-0.064215, -1.045508, -2.737277, -0.929604, 1.570796, 1.506582],accel_mss,speed_ms,0,blend_radius_m)
  movel([-0.062279, -1.041823, -2.738484, -0.932082, 1.570796, 1.508517],accel_mss,speed_ms,0,blend_radius_m)
  movel([-0.060072, -1.038263, -2.739640, -0.934486, 1.570796, 1.510725],accel_mss,speed_ms,0,blend_radius_m)
  movel([-0.052653, -1.027974, -2.742922, -0.941493, 1.570796, 1.518143],accel_mss,speed_ms,0,blend_radius_m)
  movel([-0.046893, -1.019026, -2.745708, -0.947655, 1.570796, 1.523903],accel_mss,speed_ms,0,blend_radius_m)
  movel([-0.041269, -1.009876, -2.748493, -0.954021, 1.570796, 1.529527],accel_mss,speed_ms,0,blend_radius_m)
  movel([-0.038775, -1.005705, -2.749741, -0.956944, 1.570796, 1.532021],accel_mss,speed_ms,0,blend_radius_m)
  speed_ms = 0.005
  movel([-0.038775, -0.996030, -2.744085, -0.972274, 1.570796, 1.532021],accel_mss,speed_ms,0,blend_radius_m)
  speed_ms = 0.040
  movel([-0.089816, -1.069744, -2.720244, -0.922401, 1.570796, 1.480980],accel_mss,speed_ms,0,blend_radius_m)
  speed_ms = 0.005
  movel([-0.089816, -1.079540, -2.725592, -0.907257, 1.570796, 1.480980],accel_mss,speed_ms,0,blend_radius_m)
  speed_ms = 0.025
  movel([-0.085381, -1.082583, -2.724499, -0.905307, 1.570796, 1.485415],accel_mss,speed_ms,0,blend_radius_m)
  movel([-0.083192, -1.084405, -2.723840, -0.904144, 1.570796, 1.487604],accel_mss,speed_ms,0,blend_radius_m)
  movel([-0.081191, -1.086468, -2.723091, -0.902830, 1.570796, 1.489606],accel_mss,speed_ms,0,blend_radius_m)
  movel([-0.079489, -1.088786, -2.722245, -0.901358, 1.570796, 1.491307],accel_mss,speed_ms,0,blend_radius_m)
  movel([-0.078209, -1.091381, -2.721292, -0.899717, 1.570796, 1.492587],accel_mss,speed_ms,0,blend_radius_m)
  movel([-0.077467, -1.094275, -2.720221, -0.897893, 1.570796, 1.493329],accel_mss,speed_ms,0,blend_radius_m)
  movel([-0.077335, -1.095842, -2.719639, -0.896908, 1.570796, 1.493461],accel_mss,speed_ms,0,blend_radius_m)
  movel([-0.077380, -1.097486, -2.719025, -0.895878, 1.570796, 1.493416],accel_mss,speed_ms,0,blend_radius_m)
  movel([-0.078452, -1.097177, -2.719141, -0.896071, 1.570796, 1.492345],accel_mss,speed_ms,0,blend_radius_m)
  movel([-0.079150, -1.096590, -2.719360, -0.896439, 1.570796, 1.491646],accel_mss,speed_ms,0,blend_radius_m)
  movel([-0.080624, -1.095183, -2.719884, -0.897322, 1.570796, 1.490172],accel_mss,speed_ms,0,blend_radius_m)
  movel([-0.082650, -1.094184, -2.720255, -0.897950, 1.570796, 1.488147],accel_mss,speed_ms,0,blend_radius_m)
  movel([-0.084885, -1.093461, -2.720523, -0.898405, 1.570796, 1.485911],accel_mss,speed_ms,0,blend_radius_m)
  movel([-0.087305, -1.093001, -2.720694, -0.898695, 1.570796, 1.483491],accel_mss,speed_ms,0,blend_radius_m)
  movel([-0.089883, -1.092797, -2.720769, -0.898823, 1.570796, 1.480913],accel_mss,speed_ms,0,blend_radius_m)
  movel([-0.092594, -1.092840, -2.720753, -0.898796, 1.570796, 1.478203],accel_mss,speed_ms,0,blend_radius_m)
  movel([-0.095409, -1.093121, -2.720649, -0.898619, 1.570796, 1.475387],accel_mss,speed_ms,0,blend_radius_m)
  movel([-0.098307, -1.093633, -2.720459, -0.898296, 1.570796, 1.472490],accel_mss,speed_ms,0,blend_radius_m)
  movel([-0.101256, -1.094361, -2.720189, -0.897838, 1.570796, 1.469540],accel_mss,speed_ms,0,blend_radius_m)
  movel([-0.103243, -1.095014, -2.719947, -0.897428, 1.570796, 1.467553],accel_mss,speed_ms,0,blend_radius_m)
  movel([-0.104813, -1.095730, -2.719680, -0.896978, 1.570796, 1.465983],accel_mss,speed_ms,0,blend_radius_m)
  movel([-0.105996, -1.096496, -2.719395, -0.896498, 1.570796, 1.464800],accel_mss,speed_ms,0,blend_radius_m)
  movel([-0.106828, -1.097301, -2.719094, -0.895994, 1.570796, 1.463969],accel_mss,speed_ms,0,blend_radius_m)
  movel([-0.107346, -1.098143, -2.718779, -0.895467, 1.570796, 1.463451],accel_mss,speed_ms,0,blend_radius_m)
  movel([-0.107582, -1.099011, -2.718454, -0.894924, 1.570796, 1.463214],accel_mss,speed_ms,0,blend_radius_m)
  movel([-0.107579, -1.099901, -2.718119, -0.894369, 1.570796, 1.463218],accel_mss,speed_ms,0,blend_radius_m)
  movel([-0.107365, -1.100802, -2.717780, -0.893807, 1.570796, 1.463432],accel_mss,speed_ms,0,blend_radius_m)
  movel([-0.106462, -1.102620, -2.717093, -0.892676, 1.570796, 1.464334],accel_mss,speed_ms,0,blend_radius_m)
  movel([-0.102469, -1.107720, -2.715150, -0.889519, 1.570796, 1.468328],accel_mss,speed_ms,0,blend_radius_m)
  movel([-0.105068, -1.106814, -2.715497, -0.890078, 1.570796, 1.465728],accel_mss,speed_ms,0,blend_radius_m)
  movel([-0.110164, -1.104875, -2.716237, -0.891277, 1.570796, 1.460632],accel_mss,speed_ms,0,blend_radius_m)
  movel([-0.113027, -1.104390, -2.716421, -0.891577, 1.570796, 1.457770],accel_mss,speed_ms,0,blend_radius_m)
  movel([-0.116461, -1.104328, -2.716445, -0.891616, 1.570796, 1.454335],accel_mss,speed_ms,0,blend_radius_m)
  movel([-0.120018, -1.104477, -2.716388, -0.891523, 1.570796, 1.450778],accel_mss,speed_ms,0,blend_radius_m)
  movel([-0.127213, -1.104948, -2.716209, -0.891232, 1.570796, 1.443583],accel_mss,speed_ms,0,blend_radius_m)
  movel([-0.130713, -1.105040, -2.716174, -0.891175, 1.570796, 1.440083],accel_mss,speed_ms,0,blend_radius_m)
  movel([-0.134055, -1.104883, -2.716234, -0.891272, 1.570796, 1.436742],accel_mss,speed_ms,0,blend_radius_m)
  movel([-0.137170, -1.104365, -2.716431, -0.891593, 1.570796, 1.433626],accel_mss,speed_ms,0,blend_radius_m)
  movel([-0.139995, -1.103366, -2.716810, -0.892213, 1.570796, 1.430802],accel_mss,speed_ms,0,blend_radius_m)
  movel([-0.137192, -1.107878, -2.715089, -0.889422, 1.570796, 1.433605],accel_mss,speed_ms,0,blend_radius_m)
  movel([-0.135602, -1.110055, -2.714252, -0.888082, 1.570796, 1.435194],accel_mss,speed_ms,0,blend_radius_m)
  movel([-0.133826, -1.111777, -2.713587, -0.887025, 1.570796, 1.436971],accel_mss,speed_ms,0,blend_radius_m)
  movel([-0.136672, -1.110906, -2.713924, -0.887559, 1.570796, 1.434124],accel_mss,speed_ms,0,blend_radius_m)
  movel([-0.139763, -1.110406, -2.714116, -0.887866, 1.570796, 1.431033],accel_mss,speed_ms,0,blend_radius_m)
  movel([-0.146189, -1.109788, -2.714355, -0.888246, 1.570796, 1.424608],accel_mss,speed_ms,0,blend_radius_m)
  movel([-0.148233, -1.109403, -2.714503, -0.888483, 1.570796, 1.422563],accel_mss,speed_ms,0,blend_radius_m)
  movel([-0.150068, -1.108794, -2.714737, -0.888857, 1.570796, 1.420728],accel_mss,speed_ms,0,blend_radius_m)
  movel([-0.153333, -1.107124, -2.715378, -0.889887, 1.570796, 1.417463],accel_mss,speed_ms,0,blend_radius_m)
  movel([-0.156453, -1.105243, -2.716096, -0.891049, 1.570796, 1.414344],accel_mss,speed_ms,0,blend_radius_m)
  movel([-0.159894, -1.103632, -2.716709, -0.892047, 1.570796, 1.410903],accel_mss,speed_ms,0,blend_radius_m)
  movel([-0.161112, -1.103303, -2.716834, -0.892252, 1.570796, 1.409685],accel_mss,speed_ms,0,blend_radius_m)
  movel([-0.162467, -1.103206, -2.716871, -0.892312, 1.570796, 1.408329],accel_mss,speed_ms,0,blend_radius_m)
  movel([-0.163937, -1.103492, -2.716762, -0.892134, 1.570796, 1.406859],accel_mss,speed_ms,0,blend_radius_m)
  movel([-0.164701, -1.103818, -2.716639, -0.891932, 1.570796, 1.406095],accel_mss,speed_ms,0,blend_radius_m)
  movel([-0.165483, -1.104297, -2.716457, -0.891635, 1.570796, 1.405313],accel_mss,speed_ms,0,blend_radius_m)
  movel([-0.166307, -1.104968, -2.716202, -0.891220, 1.570796, 1.404490],accel_mss,speed_ms,0,blend_radius_m)
  movel([-0.167031, -1.105732, -2.715910, -0.890747, 1.570796, 1.403765],accel_mss,speed_ms,0,blend_radius_m)
  movel([-0.168230, -1.107469, -2.715246, -0.889674, 1.570796, 1.402566],accel_mss,speed_ms,0,blend_radius_m)
  movel([-0.169139, -1.109343, -2.714526, -0.888520, 1.570796, 1.401658],accel_mss,speed_ms,0,blend_radius_m)
  movel([-0.169815, -1.111191, -2.713813, -0.887384, 1.570796, 1.400982],accel_mss,speed_ms,0,blend_radius_m)
  movel([-0.170869, -1.108921, -2.714689, -0.888779, 1.570796, 1.399927],accel_mss,speed_ms,0,blend_radius_m)
  movel([-0.172146, -1.106891, -2.715467, -0.890031, 1.570796, 1.398650],accel_mss,speed_ms,0,blend_radius_m)
  movel([-0.175130, -1.103309, -2.716832, -0.892248, 1.570796, 1.395666],accel_mss,speed_ms,0,blend_radius_m)
  movel([-0.178288, -1.099906, -2.718117, -0.894366, 1.570796, 1.392508],accel_mss,speed_ms,0,blend_radius_m)
  movel([-0.181130, -1.096124, -2.719534, -0.896731, 1.570796, 1.389666],accel_mss,speed_ms,0,blend_radius_m)
  movel([-0.181947, -1.094394, -2.720177, -0.897818, 1.570796, 1.388849],accel_mss,speed_ms,0,blend_radius_m)
  movel([-0.182498, -1.092392, -2.720919, -0.899079, 1.570796, 1.388298],accel_mss,speed_ms,0,blend_radius_m)
  movel([-0.182819, -1.090170, -2.721737, -0.900482, 1.570796, 1.387977],accel_mss,speed_ms,0,blend_radius_m)
  movel([-0.182952, -1.087790, -2.722609, -0.901990, 1.570796, 1.387845],accel_mss,speed_ms,0,blend_radius_m)
  movel([-0.182776, -1.082756, -2.724436, -0.905196, 1.570796, 1.388020],accel_mss,speed_ms,0,blend_radius_m)
  movel([-0.182269, -1.077752, -2.726231, -0.908406, 1.570796, 1.388528],accel_mss,speed_ms,0,blend_radius_m)
  speed_ms = 0.005
  movel([-0.182269, -1.067957, -2.720875, -0.923558, 1.570796, 1.388528],accel_mss,speed_ms,0,blend_radius_m)
  speed_ms = 0.040
  # Splitting Linear movement in 2 (instruction 806: MoveL 765)
  movel([-0.154336, -0.993196, -2.744917, -0.974276, 1.570796, 1.416460],accel_mss,speed_ms,0,blend_radius_m)
  movel([-0.121695, -0.908990, -2.767025, -1.036374, 1.570796, 1.449101],accel_mss,speed_ms,0,blend_radius_m)
  speed_ms = 0.005
  movel([-0.121695, -0.918267, -2.773014, -1.021108, 1.570796, 1.449101],accel_mss,speed_ms,0,blend_radius_m)
  speed_ms = 0.025
  movel([-0.123729, -0.920795, -2.772414, -1.019180, 1.570796, 1.447067],accel_mss,speed_ms,0,blend_radius_m)
  movel([-0.123869, -0.921211, -2.772315, -1.018863, 1.570796, 1.446928],accel_mss,speed_ms,0,blend_radius_m)
  movel([-0.123677, -0.921670, -2.772206, -1.018514, 1.570796, 1.447119],accel_mss,speed_ms,0,blend_radius_m)
  movel([-0.122387, -0.922727, -2.771953, -1.017709, 1.570796, 1.448409],accel_mss,speed_ms,0,blend_radius_m)
  movel([-0.116786, -0.925304, -2.771334, -1.015751, 1.570796, 1.454011],accel_mss,speed_ms,0,blend_radius_m)
  movel([-0.108296, -0.928361, -2.770594, -1.013434, 1.570796, 1.462501],accel_mss,speed_ms,0,blend_radius_m)
  movel([-0.098262, -0.931706, -2.769778, -1.010905, 1.570796, 1.472535],accel_mss,speed_ms,0,blend_radius_m)
  movel([-0.078691, -0.938178, -2.768177, -1.006034, 1.570796, 1.492105],accel_mss,speed_ms,0,blend_radius_m)
  movel([-0.067694, -0.941754, -2.767280, -1.003355, 1.570796, 1.503103],accel_mss,speed_ms,0,blend_radius_m)
  movel([-0.066628, -0.941922, -2.767238, -1.003229, 1.570796, 1.504168],accel_mss,speed_ms,0,blend_radius_m)
  movel([-0.065426, -0.941835, -2.767260, -1.003294, 1.570796, 1.505370],accel_mss,speed_ms,0,blend_radius_m)
  movel([-0.064169, -0.941340, -2.767384, -1.003664, 1.570796, 1.506628],accel_mss,speed_ms,0,blend_radius_m)
  movel([-0.063539, -0.940894, -2.767497, -1.003998, 1.570796, 1.507257],accel_mss,speed_ms,0,blend_radius_m)
  movel([-0.062925, -0.940286, -2.767649, -1.004453, 1.570796, 1.507871],accel_mss,speed_ms,0,blend_radius_m)
  movel([-0.062039, -0.938976, -2.767977, -1.005435, 1.570796, 1.508758],accel_mss,speed_ms,0,blend_radius_m)
  movel([-0.061407, -0.937605, -2.768320, -1.006464, 1.570796, 1.509389],accel_mss,speed_ms,0,blend_radius_m)
  movel([-0.058516, -0.929995, -2.770196, -1.012198, 1.570796, 1.512280],accel_mss,speed_ms,0,blend_radius_m)
  movel([-0.056125, -0.922455, -2.772018, -1.017916, 1.570796, 1.514671],accel_mss,speed_ms,0,blend_radius_m)
  movel([-0.054216, -0.915024, -2.773777, -1.023587, 1.570796, 1.516580],accel_mss,speed_ms,0,blend_radius_m)
  movel([-0.052750, -0.907727, -2.775471, -1.029191, 1.570796, 1.518046],accel_mss,speed_ms,0,blend_radius_m)
  movel([-0.051705, -0.900594, -2.777094, -1.034701, 1.570796, 1.519091],accel_mss,speed_ms,0,blend_radius_m)
  movel([-0.051044, -0.893651, -2.778643, -1.040095, 1.570796, 1.519752],accel_mss,speed_ms,0,blend_radius_m)
  movel([-0.050737, -0.886930, -2.780115, -1.045344, 1.570796, 1.520059],accel_mss,speed_ms,0,blend_radius_m)
  movel([-0.050750, -0.880465, -2.781505, -1.050419, 1.570796, 1.520046],accel_mss,speed_ms,0,blend_radius_m)
  movel([-0.050960, -0.877664, -2.782100, -1.052626, 1.570796, 1.519836],accel_mss,speed_ms,0,blend_radius_m)
  movel([-0.051433, -0.875241, -2.782610, -1.054538, 1.570796, 1.519363],accel_mss,speed_ms,0,blend_radius_m)
  movel([-0.052166, -0.873195, -2.783038, -1.056156, 1.570796, 1.518631],accel_mss,speed_ms,0,blend_radius_m)
  movel([-0.053142, -0.871512, -2.783389, -1.057488, 1.570796, 1.517655],accel_mss,speed_ms,0,blend_radius_m)
  movel([-0.054358, -0.870191, -2.783662, -1.058535, 1.570796, 1.516439],accel_mss,speed_ms,0,blend_radius_m)
  movel([-0.055805, -0.869228, -2.783861, -1.059299, 1.570796, 1.514992],accel_mss,speed_ms,0,blend_radius_m)
  movel([-0.057470, -0.868603, -2.783990, -1.059795, 1.570796, 1.513326],accel_mss,speed_ms,0,blend_radius_m)
  movel([-0.059349, -0.868314, -2.784050, -1.060025, 1.570796, 1.511448],accel_mss,speed_ms,0,blend_radius_m)
  movel([-0.061426, -0.868351, -2.784042, -1.059996, 1.570796, 1.509370],accel_mss,speed_ms,0,blend_radius_m)
  movel([-0.063692, -0.868703, -2.783970, -1.059716, 1.570796, 1.507104],accel_mss,speed_ms,0,blend_radius_m)
  movel([-0.066142, -0.869359, -2.783834, -1.059195, 1.570796, 1.504655],accel_mss,speed_ms,0,blend_radius_m)
  movel([-0.068755, -0.870309, -2.783638, -1.058442, 1.570796, 1.502042],accel_mss,speed_ms,0,blend_radius_m)
  movel([-0.074446, -0.873048, -2.783069, -1.056272, 1.570796, 1.496350],accel_mss,speed_ms,0,blend_radius_m)
  movel([-0.080671, -0.876818, -2.782278, -1.053293, 1.570796, 1.490125],accel_mss,speed_ms,0,blend_radius_m)
  movel([-0.086258, -0.880831, -2.781427, -1.050131, 1.570796, 1.484538],accel_mss,speed_ms,0,blend_radius_m)
  movel([-0.091716, -0.885353, -2.780457, -1.046580, 1.570796, 1.479080],accel_mss,speed_ms,0,blend_radius_m)
  movel([-0.097048, -0.890304, -2.779380, -1.042705, 1.570796, 1.473748],accel_mss,speed_ms,0,blend_radius_m)
  movel([-0.102248, -0.895586, -2.778215, -1.038589, 1.570796, 1.468548],accel_mss,speed_ms,0,blend_radius_m)
  movel([-0.107307, -0.901104, -2.776979, -1.034306, 1.570796, 1.463490],accel_mss,speed_ms,0,blend_radius_m)
  movel([-0.112236, -0.906780, -2.775688, -1.029921, 1.570796, 1.458561],accel_mss,speed_ms,0,blend_radius_m)
  movel([-0.121695, -0.918267, -2.773014, -1.021108, 1.570796, 1.449101],accel_mss,speed_ms,0,blend_radius_m)
  movel([-0.123729, -0.920795, -2.772414, -1.019180, 1.570796, 1.447067],accel_mss,speed_ms,0,blend_radius_m)
  movel([-0.123869, -0.921211, -2.772315, -1.018863, 1.570796, 1.446928],accel_mss,speed_ms,0,blend_radius_m)
  movel([-0.123677, -0.921670, -2.772206, -1.018514, 1.570796, 1.447119],accel_mss,speed_ms,0,blend_radius_m)
  movel([-0.123269, -0.922006, -2.772125, -1.018258, 1.570796, 1.447527],accel_mss,speed_ms,0,blend_radius_m)
  speed_ms = 0.005
  movel([-0.123269, -0.912705, -2.766150, -1.033534, 1.570796, 1.447527],accel_mss,speed_ms,0,blend_radius_m)
  speed_ms = 0.040
  movel([-0.141809, -0.890212, -2.771314, -1.050863, 1.570796, 1.428988],accel_mss,speed_ms,0,blend_radius_m)
  speed_ms = 0.005
  movel([-0.141809, -0.899367, -2.777370, -1.035652, 1.570796, 1.428988],accel_mss,speed_ms,0,blend_radius_m)
  speed_ms = 0.025
  movel([-0.142140, -0.896959, -2.777909, -1.037521, 1.570796, 1.428656],accel_mss,speed_ms,0,blend_radius_m)
  movel([-0.142908, -0.894918, -2.778363, -1.039108, 1.570796, 1.427888],accel_mss,speed_ms,0,blend_radius_m)
  movel([-0.144096, -0.893298, -2.778721, -1.040370, 1.570796, 1.426701],accel_mss,speed_ms,0,blend_radius_m)
  movel([-0.145674, -0.892135, -2.778978, -1.041276, 1.570796, 1.425122],accel_mss,speed_ms,0,blend_radius_m)
  movel([-0.150413, -0.890446, -2.779349, -1.042594, 1.570796, 1.420383],accel_mss,speed_ms,0,blend_radius_m)
  movel([-0.151583, -0.889732, -2.779505, -1.043152, 1.570796, 1.419213],accel_mss,speed_ms,0,blend_radius_m)
  movel([-0.152432, -0.888798, -2.779709, -1.043882, 1.570796, 1.418365],accel_mss,speed_ms,0,blend_radius_m)
  movel([-0.152803, -0.887599, -2.779970, -1.044820, 1.570796, 1.417993],accel_mss,speed_ms,0,blend_radius_m)
  movel([-0.152536, -0.886075, -2.780300, -1.046014, 1.570796, 1.418260],accel_mss,speed_ms,0,blend_radius_m)
  movel([-0.151543, -0.884128, -2.780721, -1.047541, 1.570796, 1.419254],accel_mss,speed_ms,0,blend_radius_m)
  movel([-0.150265, -0.882614, -2.781046, -1.048729, 1.570796, 1.420531],accel_mss,speed_ms,0,blend_radius_m)
  movel([-0.148786, -0.881480, -2.781288, -1.049620, 1.570796, 1.422010],accel_mss,speed_ms,0,blend_radius_m)
  movel([-0.147199, -0.880675, -2.781460, -1.050254, 1.570796, 1.423597],accel_mss,speed_ms,0,blend_radius_m)
  movel([-0.144077, -0.879854, -2.781635, -1.050900, 1.570796, 1.426719],accel_mss,speed_ms,0,blend_radius_m)
  movel([-0.141608, -0.879725, -2.781663, -1.051002, 1.570796, 1.429189],accel_mss,speed_ms,0,blend_radius_m)
  movel([-0.142716, -0.877240, -2.782189, -1.052960, 1.570796, 1.428081],accel_mss,speed_ms,0,blend_radius_m)
  movel([-0.144331, -0.875361, -2.782585, -1.054443, 1.570796, 1.426465],accel_mss,speed_ms,0,blend_radius_m)
  movel([-0.148487, -0.872677, -2.783146, -1.056566, 1.570796, 1.422309],accel_mss,speed_ms,0,blend_radius_m)
  movel([-0.152861, -0.870136, -2.783674, -1.058579, 1.570796, 1.417935],accel_mss,speed_ms,0,blend_radius_m)
  movel([-0.154755, -0.868431, -2.784026, -1.059932, 1.570796, 1.416041],accel_mss,speed_ms,0,blend_radius_m)
  movel([-0.156241, -0.866167, -2.784491, -1.061731, 1.570796, 1.414555],accel_mss,speed_ms,0,blend_radius_m)
  movel([-0.156900, -0.864453, -2.784840, -1.063095, 1.570796, 1.413896],accel_mss,speed_ms,0,blend_radius_m)
  movel([-0.157213, -0.862866, -2.785163, -1.064360, 1.570796, 1.413584],accel_mss,speed_ms,0,blend_radius_m)
  movel([-0.157211, -0.861410, -2.785457, -1.065522, 1.570796, 1.413585],accel_mss,speed_ms,0,blend_radius_m)
  movel([-0.156924, -0.860093, -2.785723, -1.066574, 1.570796, 1.413873],accel_mss,speed_ms,0,blend_radius_m)
  movel([-0.156395, -0.858928, -2.785956, -1.067504, 1.570796, 1.414402],accel_mss,speed_ms,0,blend_radius_m)
  movel([-0.155651, -0.857912, -2.786160, -1.068317, 1.570796, 1.415145],accel_mss,speed_ms,0,blend_radius_m)
  movel([-0.154736, -0.857061, -2.786330, -1.068999, 1.570796, 1.416060],accel_mss,speed_ms,0,blend_radius_m)
  movel([-0.153677, -0.856378, -2.786466, -1.069545, 1.570796, 1.417119],accel_mss,speed_ms,0,blend_radius_m)
  movel([-0.152514, -0.855873, -2.786566, -1.069950, 1.570796, 1.418282],accel_mss,speed_ms,0,blend_radius_m)
  movel([-0.151289, -0.855558, -2.786629, -1.070202, 1.570796, 1.419507],accel_mss,speed_ms,0,blend_radius_m)
  movel([-0.148777, -0.855513, -2.786638, -1.070238, 1.570796, 1.422019],accel_mss,speed_ms,0,blend_radius_m)
  movel([-0.146432, -0.856297, -2.786482, -1.069610, 1.570796, 1.424365],accel_mss,speed_ms,0,blend_radius_m)
  movel([-0.144538, -0.857966, -2.786149, -1.068274, 1.570796, 1.426258],accel_mss,speed_ms,0,blend_radius_m)
  movel([-0.144291, -0.854919, -2.786755, -1.070714, 1.570796, 1.426505],accel_mss,speed_ms,0,blend_radius_m)
  movel([-0.144419, -0.852292, -2.787274, -1.072823, 1.570796, 1.426377],accel_mss,speed_ms,0,blend_radius_m)
  movel([-0.144844, -0.849994, -2.787724, -1.074671, 1.570796, 1.425952],accel_mss,speed_ms,0,blend_radius_m)
  movel([-0.147033, -0.843965, -2.788892, -1.079533, 1.570796, 1.423764],accel_mss,speed_ms,0,blend_radius_m)
  movel([-0.148397, -0.839580, -2.789728, -1.083081, 1.570796, 1.422399],accel_mss,speed_ms,0,blend_radius_m)
  movel([-0.148692, -0.837536, -2.790114, -1.084739, 1.570796, 1.422104],accel_mss,speed_ms,0,blend_radius_m)
  movel([-0.148704, -0.835573, -2.790483, -1.086333, 1.570796, 1.422092],accel_mss,speed_ms,0,blend_radius_m)
  movel([-0.148469, -0.833724, -2.790828, -1.087837, 1.570796, 1.422328],accel_mss,speed_ms,0,blend_radius_m)
  movel([-0.148012, -0.832008, -2.791147, -1.089234, 1.570796, 1.422784],accel_mss,speed_ms,0,blend_radius_m)
  movel([-0.147373, -0.830451, -2.791435, -1.090503, 1.570796, 1.423424],accel_mss,speed_ms,0,blend_radius_m)
  movel([-0.146578, -0.829074, -2.791688, -1.091627, 1.570796, 1.424218],accel_mss,speed_ms,0,blend_radius_m)
  movel([-0.145663, -0.827902, -2.791903, -1.092584, 1.570796, 1.425134],accel_mss,speed_ms,0,blend_radius_m)
  movel([-0.144659, -0.826962, -2.792075, -1.093352, 1.570796, 1.426137],accel_mss,speed_ms,0,blend_radius_m)
  movel([-0.143601, -0.826279, -2.792200, -1.093910, 1.570796, 1.427195],accel_mss,speed_ms,0,blend_radius_m)
  movel([-0.142525, -0.825876, -2.792273, -1.094240, 1.570796, 1.428271],accel_mss,speed_ms,0,blend_radius_m)
  movel([-0.141459, -0.825775, -2.792292, -1.094323, 1.570796, 1.429337],accel_mss,speed_ms,0,blend_radius_m)
  movel([-0.140438, -0.826004, -2.792250, -1.094135, 1.570796, 1.430358],accel_mss,speed_ms,0,blend_radius_m)
  movel([-0.139501, -0.826588, -2.792143, -1.093657, 1.570796, 1.431295],accel_mss,speed_ms,0,blend_radius_m)
  movel([-0.138678, -0.827549, -2.791968, -1.092872, 1.570796, 1.432119],accel_mss,speed_ms,0,blend_radius_m)
  movel([-0.138001, -0.828909, -2.791719, -1.091762, 1.570796, 1.432795],accel_mss,speed_ms,0,blend_radius_m)
  movel([-0.137501, -0.830682, -2.791392, -1.090315, 1.570796, 1.433296],accel_mss,speed_ms,0,blend_radius_m)
  movel([-0.136094, -0.827442, -2.791987, -1.092959, 1.570796, 1.434702],accel_mss,speed_ms,0,blend_radius_m)
  movel([-0.135009, -0.824327, -2.792554, -1.095508, 1.570796, 1.435788],accel_mss,speed_ms,0,blend_radius_m)
  movel([-0.134183, -0.821312, -2.793098, -1.097979, 1.570796, 1.436613],accel_mss,speed_ms,0,blend_radius_m)
  movel([-0.133548, -0.818369, -2.793624, -1.100396, 1.570796, 1.437248],accel_mss,speed_ms,0,blend_radius_m)
  movel([-0.131530, -0.806779, -2.795651, -1.109959, 1.570796, 1.439266],accel_mss,speed_ms,0,blend_radius_m)
  movel([-0.130668, -0.802430, -2.796393, -1.113566, 1.570796, 1.440128],accel_mss,speed_ms,0,blend_radius_m)
  movel([-0.129218, -0.797065, -2.797295, -1.118029, 1.570796, 1.441578],accel_mss,speed_ms,0,blend_radius_m)
  movel([-0.128102, -0.794324, -2.797750, -1.120315, 1.570796, 1.442695],accel_mss,speed_ms,0,blend_radius_m)
  movel([-0.126634, -0.791725, -2.798178, -1.122485, 1.570796, 1.444162],accel_mss,speed_ms,0,blend_radius_m)
  movel([-0.125742, -0.790517, -2.798376, -1.123496, 1.570796, 1.445055],accel_mss,speed_ms,0,blend_radius_m)
